(* IEC 61131-3 sources: daoli-st-library/DL_MathData (part 14) *)

(* ---- FC_DL_GearModuleFromCpCalc.st ---- *)
(*
  DL Factory R88 | FC_DL_GearModuleFromCpCalc
  功能：由圆周节 Cp 反算齿轮模数 m=Cp/π，并校验模数是否落在 [min,max] 允许区间
  开源溯源：无（clean-room 自研，依据公开工艺公式 圆周节-模数关系 m=Cp/π，许可证=MIT，借鉴点=公式结构）
  规则：R1-R16 全遵守；R88 简单件标量形（纯标量入参出参，无循环体、无方法、无属性、无数组）
*)
FUNCTION FC_DL_GearModuleFromCpCalc : REAL
VAR_INPUT
    fCpMm : REAL := 12.56637; // 圆周节 Cp（分度圆上相邻同侧齿廓的弧长） [mm] / circular pitch [mm]
    fModuleMin : REAL := 1.0; // 模数允许下限 [mm] / lower allowed module [mm]
    fModuleMax : REAL := 10.0; // 模数允许上限 [mm] / upper allowed module [mm]
END_VAR
VAR_OUTPUT
    fModuleMm : REAL; // 反算模数 m [mm] / back calculated module [mm]
    xInRange : BOOL; // TRUE=模数落在允许区间 [-] / TRUE when module inside the band [-]
END_VAR
VAR
    fPiC : REAL; // 圆周率常数（REAL 精度装入，避免长字面量截断） [-] / pi constant in REAL precision [-]
END_VAR

// 段 1｜出口预置
FC_DL_GearModuleFromCpCalc := -1.0; // 哨兵返回 -1（无效） [-] / sentinel return -1, invalid [-]
fModuleMm := 0.0; // 模数出口预置零 [mm] / module output preset zero [mm]
xInRange := FALSE; // 区间位预置 FALSE（未判定前不认合格） [-] / in-range preset false [-]
fPiC := 3.14159265; // π 常数装入，无量纲 [-] / load the pi constant, dimensionless [-]

// 段 2｜非有限拦截 + 域闸
IF NOT (fCpMm > -1.0E30 AND fCpMm < 1.0E30) OR NOT (fModuleMin > -1.0E30 AND fModuleMin < 1.0E30) OR NOT (fModuleMax > -1.0E30 AND fModuleMax < 1.0E30) THEN
    RETURN; // 三入参任一非有限（NaN/±Inf）即拒算 [-] / any non finite input rejected [-]
END_IF
IF fCpMm < 1.0E-9 THEN
    RETURN; // 周节正域闸：分母 π 恒正，此处拦非正的周节输入 [mm] / positive circular pitch gate [mm]
END_IF
IF fModuleMin < 1.0E-9 OR fModuleMax <= fModuleMin THEN
    RETURN; // 区间自洽闸：下限须为正、上限须严格大于下限 [mm] / band consistency gate [mm]
END_IF

// 段 3｜计算
fModuleMm := fCpMm / fPiC; // mm ÷ 无量纲 = mm，即 m=Cp/π / [mm] / [-] = [mm], m = Cp / pi

// 段 4｜判定与饱和
IF NOT (fModuleMm > -1.0E30 AND fModuleMm < 1.0E30) THEN
    RETURN; // 商结果非有限再拦一次，防溢出成 Inf [-] / re-check the quotient for finiteness [-]
END_IF
xInRange := (fModuleMm >= fModuleMin) AND (fModuleMm <= fModuleMax); // 双侧闭区间直比（含边界） [mm] / closed two sided band compare [mm]

// 段 5｜出口自检
IF fModuleMm < 1.0E-9 THEN
    RETURN; // 出口自检：模数须为正，否则退回哨兵 [mm] / exit self-check, module must be positive [mm]
END_IF
FC_DL_GearModuleFromCpCalc := fModuleMm; // 返回反算模数 [mm] / return the back calculated module [mm]
END_FUNCTION

(* ---- FC_DL_GearRootCircleCalc.st ---- *)
(*
  DL Factory R88 | FC_DL_GearRootCircleCalc
  功能：由模数/齿数算齿根圆直径 df=m(z-2.5)（等价 d-2hf，hf=1.25m），齿数域闸 z>=8
  开源溯源：无（clean-room 自研，依据公开工艺公式 齿根圆直径式 df=m(z-2.5)，许可证=MIT，借鉴点=公式结构）
  规则：R1-R16 全遵守；R88 简单件标量形（纯标量入参出参，无循环体、无方法、无属性、无数组）
*)
FUNCTION FC_DL_GearRootCircleCalc : REAL
VAR_INPUT
    fModuleMm : REAL := 3.0; // 模数 m [mm] / module [mm]
    nTeeth : DINT := 20; // 齿数 z，域闸 z>=8 防齿根自交 [枚] / tooth count, gated at 8 or more [-]
    fDedFactor : REAL := 1.25; // 齿根高系数 hf*=1.25，使 2hf*=2.5 与公式一致 [-] / dedendum coefficient [-]
END_VAR
VAR_OUTPUT
    fDfMm : REAL; // 齿根圆直径 df [mm] / root circle diameter [mm]
    fDedendumMm : REAL; // 齿根高 hf=hf*·m [mm] / dedendum height [mm]
END_VAR
VAR
    fTeeth : REAL; // 齿数实数化结果 [-] / tooth count converted to REAL [-]
    fPitchDiaMm : REAL; // 分度圆直径 d=m·z [mm] / pitch circle diameter [mm]
END_VAR

// 段 1｜出口预置
FC_DL_GearRootCircleCalc := -1.0; // 哨兵返回 -1（无效） [-] / sentinel return -1, invalid [-]
fDfMm := 0.0; // 齿根圆直径预置零 [mm] / root diameter preset zero [mm]
fDedendumMm := 0.0; // 齿根高预置零 [mm] / dedendum preset zero [mm]
fTeeth := 0.0; // 齿数实数预置零 [-] / real teeth preset zero [-]
fPitchDiaMm := 0.0; // 分度圆直径预置零 [mm] / pitch diameter preset zero [mm]

// 段 2｜非有限拦截 + 域闸
IF NOT (fModuleMm > -1.0E30 AND fModuleMm < 1.0E30) OR NOT (fDedFactor > -1.0E30 AND fDedFactor < 1.0E30) THEN
    RETURN; // 模数/齿根高系数任一非有限即拒算 [-] / any non finite input rejected [-]
END_IF
IF fModuleMm < 1.0E-9 THEN
    RETURN; // 模数正域闸 [mm] / positive module gate [mm]
END_IF
IF fDedFactor < 0.8 OR fDedFactor > 1.6 THEN
    RETURN; // 齿根高系数工程域闸（0.8~1.6，标准 1.25） [-] / dedendum coefficient domain gate [-]
END_IF
IF nTeeth < 8 THEN
    RETURN; // 齿数域闸 z>=8：低于 8 齿时齿根圆退化、公式失真 [枚] / root circle degenerates below 8 teeth [-]
END_IF

// 段 3｜计算
fTeeth := DINT_TO_REAL(nTeeth); // DINT→REAL 标准转换函数（R10） [-] / standard conversion function (R10) [-]
fDedendumMm := fDedFactor * fModuleMm; // 无量纲 × mm = mm，hf=hf*·m / [-] × [mm] = [mm]
fPitchDiaMm := fModuleMm * fTeeth; // mm × 无量纲 = mm，d=m·z / [mm] × [-] = [mm]
fDfMm := fPitchDiaMm - 2.0 * fDedendumMm; // mm - mm = mm，df=d-2hf=m(z-2.5) / [mm]

// 段 4｜判定与饱和
IF fDfMm <= 0.0 THEN
    RETURN; // 结果闸：齿根圆直径必须为正，否则齿形无意义 [mm] / root diameter must be positive [mm]
END_IF
IF fDfMm >= fPitchDiaMm THEN
    RETURN; // 结构自洽闸：齿根圆必须小于分度圆 [mm] / structural check df < d [mm]
END_IF

// 段 5｜出口自检
IF NOT (fDfMm > -1.0E30 AND fDfMm < 1.0E30) THEN
    RETURN; // 出口自检：结果非有限即退回哨兵 [mm] / exit self-check on finiteness [mm]
END_IF
FC_DL_GearRootCircleCalc := fDfMm; // 返回齿根圆直径 [mm] / return the root circle diameter [mm]
END_FUNCTION

(* ---- FC_DL_GearSpanMeasurementCalc.st ---- *)
(*
  DL Factory R88 | FC_DL_GearSpanMeasurementCalc
  功能：由模数/齿数/压力角算跨 k 齿公法线长度 Wk=m·cosα·[π(k-0.5)+z·invα]
  开源溯源：无（clean-room 自研，依据公开工艺公式 跨齿公法线长度式，许可证=MIT，借鉴点=公式结构）
  规则：R1-R16 全遵守；R88 简单件标量形（纯标量入参出参，无循环体、无方法、无属性、无数组）
*)
FUNCTION FC_DL_GearSpanMeasurementCalc : REAL
VAR_INPUT
    fModuleMm : REAL := 3.0; // 模数 m [mm] / module [mm]
    nTeeth : DINT := 20; // 齿数 z（整数入参，无 NaN 可能，需 z>=5） [枚] / tooth count [-]
    fPressureDeg : REAL := 20.0; // 分度圆压力角 α（度制，域闸 10~30） [°] / pressure angle in degrees [-]
END_VAR
VAR_OUTPUT
    fWkMm : REAL; // 跨 k 齿公法线长度 Wk [mm] / span measurement over k teeth [mm]
    nSpanTeeth : REAL; // 跨齿数 k（REAL 承载的近似整数） [枚] / number of spanned teeth as a real [-]
END_VAR
VAR
    fTeeth : REAL; // 齿数实数化结果 [-] / tooth count converted to REAL [-]
    fAlphaRad : REAL; // 压力角弧度值 [rad] / pressure angle in radians [rad]
    fInvAlpha : REAL; // 渐开线函数 invα=tanα-α(rad) [rad] / involute function [rad]
    fK : REAL; // 取整后的跨齿数 [枚] / truncated span count [-]
    fCosAlpha : REAL; // 压力角余弦 [-] / cosine of the pressure angle [-]
END_VAR

// 段 1｜出口预置
FC_DL_GearSpanMeasurementCalc := -1.0; // 哨兵返回 -1（无效） [-] / sentinel return -1, invalid [-]
fWkMm := 0.0; // 公法线长度预置零 [mm] / span measurement preset zero [mm]
nSpanTeeth := 0.0; // 跨齿数预置零 [枚] / span teeth preset zero [-]

// 段 2｜非有限拦截 + 域闸
IF NOT (fModuleMm > -1.0E30 AND fModuleMm < 1.0E30) OR NOT (fPressureDeg > -1.0E30 AND fPressureDeg < 1.0E30) THEN
    RETURN; // 模数/压力角任一非有限即拒算 [-] / any non finite input rejected [-]
END_IF
IF fModuleMm < 1.0E-9 THEN
    RETURN; // 模数正域闸 [mm] / positive module gate [mm]
END_IF
IF fPressureDeg <= 10.0 OR fPressureDeg >= 30.0 THEN
    RETURN; // 压力角开区间域闸 (10°,30°)，防 invα 与 k 估算同时失真 [°] / open interval gate on alpha [deg]
END_IF
IF nTeeth < 5 THEN
    RETURN; // 齿数下限闸：z<5 时跨齿数估算式不成立 [枚] / span formula invalid below 5 teeth [-]
END_IF

// 段 3｜计算
fTeeth := DINT_TO_REAL(nTeeth); // DINT→REAL 标准转换函数（R10 禁构造函数式） [-] / standard conversion (R10) [-]
fAlphaRad := fPressureDeg * 0.0174532925; // 度 × (π/180) = rad，换算常数 0.0174532925 [rad] / degrees to radians [rad]
fInvAlpha := TAN(fAlphaRad) - fAlphaRad; // tanα-α 均取弧度，结果弧度制 [rad] / involute function in radians [rad]
fCosAlpha := COS(fAlphaRad); // 无量纲 [-] / dimensionless cosine [-]
// 跨齿数估算：k = ROUND(z·α/180 + 0.5)（标准表 z=20/α=20°→3、z=30→4、z=40→5）；正数下 ROUND 等价 TRUNC(x+1)
fK := TRUNC(fTeeth * fPressureDeg / 180.0 + 1.0); // 数学等价 ROUND(z·α/180+0.5)（R88 修复：原式少 1 齿） [枚] / span count [-]
IF fK < 1.0 THEN
    fK := 1.0; // 饱和：跨齿数至少 1，防 k<=0 使公式失效 [枚] / saturate the span count at one [-]
END_IF
nSpanTeeth := fK; // 跨齿数出口（REAL 承载近似整数） [枚] / export span teeth as a real [-]
fWkMm := fModuleMm * fCosAlpha * (3.14159265 * (fK - 0.5) + fTeeth * fInvAlpha); // mm × [-] × [-] = mm，Wk [mm] / span measurement [mm]
IF fWkMm <= 0.0 THEN
    RETURN; // 结果闸：公法线长度必须为正，否则跨齿数取值失败 [mm] / span length must be positive [mm]
END_IF

// 段 4｜判定与饱和
IF NOT (fWkMm > -1.0E30 AND fWkMm < 1.0E30) THEN
    RETURN; // 结果非有限再拦一次 [-] / re-check the result for finiteness [-]
END_IF

// 段 5｜出口自检
IF nSpanTeeth < 1.0 OR nSpanTeeth >= fTeeth THEN
    RETURN; // 出口自检：跨齿数须在 [1,z) 内，否则出口不自洽 [枚] / span count must lie in [1,z) [-]
END_IF
FC_DL_GearSpanMeasurementCalc := fWkMm; // 返回跨 k 齿公法线长度 [mm] / return the span measurement [mm]
END_FUNCTION

(* ---- FC_DL_GearToothThicknessCalc.st ---- *)
(*
  DL Factory R88 | FC_DL_GearToothThicknessCalc
  功能：由模数/齿数算分度圆弦齿厚 s=m·z·sin(π/(2z))，并给出弧齿厚 πm/2 参考值，齿数域闸 z>=6
  开源溯源：无（clean-room 自研，依据公开工艺公式 分度圆弦齿厚式 s=d·sin(π/2z)，许可证=MIT，借鉴点=公式结构）
  规则：R1-R16 全遵守；R88 简单件标量形（纯标量入参出参，无循环体、无方法、无属性、无数组）
*)
FUNCTION FC_DL_GearToothThicknessCalc : REAL
VAR_INPUT
    fModuleMm : REAL := 3.0; // 模数 m [mm] / module [mm]
    nTeeth : DINT := 20; // 齿数 z，域闸 z>=6 [枚] / tooth count, gated at 6 or more [-]
    fHalfAngleMaxRad : REAL := 1.5; // 半齿角上限保护（π/(2z) 须小于此值，防高齿数误用） [rad] / half tooth angle ceiling [rad]
END_VAR
VAR_OUTPUT
    fChordThkMm : REAL; // 分度圆弦齿厚 s [mm] / chordal tooth thickness [mm]
    fArcThkMm : REAL; // 分度圆弧齿厚 πm/2（参考值） [mm] / circular tooth thickness reference [mm]
END_VAR
VAR
    fTeeth : REAL; // 齿数实数化结果 [-] / tooth count converted to REAL [-]
    fHalfAngleRad : REAL; // 半齿角 π/(2z) [rad] / half tooth angle [rad]
    fDenomTeeth : REAL; // 半齿角分母 2z（除零判据） [枚] / half angle denominator [-]
END_VAR

// 段 1｜出口预置
FC_DL_GearToothThicknessCalc := -1.0; // 哨兵返回 -1（无效） [-] / sentinel return -1, invalid [-]
fChordThkMm := 0.0; // 弦齿厚预置零 [mm] / chordal thickness preset zero [mm]
fArcThkMm := 0.0; // 弧齿厚预置零 [mm] / circular thickness preset zero [mm]
fTeeth := 0.0; // 齿数实数预置零 [-] / real teeth preset zero [-]
fHalfAngleRad := 0.0; // 半齿角预置零 [rad] / half angle preset zero [rad]
fDenomTeeth := 0.0; // 分母预置零 [枚] / denominator preset zero [-]

// 段 2｜非有限拦截 + 域闸
IF NOT (fModuleMm > -1.0E30 AND fModuleMm < 1.0E30) OR NOT (fHalfAngleMaxRad > -1.0E30 AND fHalfAngleMaxRad < 1.0E30) THEN
    RETURN; // 模数/保护限任一非有限即拒算 [-] / any non finite input rejected [-]
END_IF
IF fModuleMm < 1.0E-9 THEN
    RETURN; // 模数正域闸 [mm] / positive module gate [mm]
END_IF
IF fHalfAngleMaxRad <= 0.0 THEN
    RETURN; // 保护限正域闸：须为正，否则后面判据失效 [rad] / positive ceiling gate [rad]
END_IF
IF nTeeth < 6 THEN
    RETURN; // 齿数域闸 z>=6：齿数过低时弦齿厚式与齿形均失真 [枚] / tooth count gate for the chord formula [-]
END_IF

// 段 3｜计算
fTeeth := DINT_TO_REAL(nTeeth); // DINT→REAL 标准转换函数（R10） [-] / standard conversion function (R10) [-]
fDenomTeeth := 2.0 * fTeeth; // 无量纲 × 无量纲 = 无量纲，即 2z [-] / the 2z denominator [-]
IF fDenomTeeth < 1.0E-9 THEN
    RETURN; // 除法前分母闸：2z 必须大于 1E-9 才可作除数 [-] / denominator gate before the division [-]
END_IF
fHalfAngleRad := 3.14159265 / fDenomTeeth; // 无量纲 ÷ 无量纲 = rad，π/(2z) [rad] / half tooth angle [rad]
IF fHalfAngleRad >= fHalfAngleMaxRad THEN
    RETURN; // 半齿角上限闸：超出说明齿数或输入落入误用区间 [rad] / half angle ceiling check [rad]
END_IF
fChordThkMm := fModuleMm * fTeeth * SIN(fHalfAngleRad); // mm × [-] × [-] = mm，s=m·z·sin(π/2z) / [mm]
fArcThkMm := 3.14159265 * fModuleMm * 0.5; // 无量纲 × mm × 0.5 = mm，πm/2（以乘 0.5 替除 2） / [mm]

// 段 4｜判定与饱和
IF fChordThkMm <= 0.0 OR fChordThkMm >= fArcThkMm THEN
    RETURN; // 结构自洽闸：弦齿厚须为正且小于弧齿厚 [mm] / chord thickness must lie in (0, arc) [mm]
END_IF

// 段 5｜出口自检
IF NOT (fChordThkMm > -1.0E30 AND fChordThkMm < 1.0E30) THEN
    RETURN; // 出口自检：结果非有限即退回哨兵 [mm] / exit self-check on finiteness [mm]
END_IF
FC_DL_GearToothThicknessCalc := fChordThkMm; // 返回分度圆弦齿厚 [mm] / return the chordal tooth thickness [mm]
END_FUNCTION

(* ---- FC_DL_GeoBBoxFromPtsFixed.st ---- *)
(*==============================================================================
 * 组件名称 : FC_DL_GeoBBoxFromPtsFixed ｜ 子库 : DL_MathData ｜ v1.0.0 ｜ 2026-11-24
 * 平台     : CODESYS 3.5 / TwinCAT 3 / InoProShop / Machine Expert（纯 IEC，无厂商库）
 * 功能简介 : 定长点列的轴对齐包围盒（BBox）。出参四个极值，用于视觉 ROI 自动贴合、
 *            轨迹占位评估、图形显示自适应缩放。
 * 契约     : 成功返回 TRUE 并写出 fMinX / fMaxX / fMinY / fMaxY；nCnt < 1 时返回 FALSE、
 *            bError := TRUE、四出参置 0；nCnt > 10 时钳到 10 继续（钳位为确定结论）。
 *            数组定长 ARRAY[1..10]，禁变长形参（R17）。
 * 依赖     : 无 DL_ 内部依赖（R16 自足实现），无标准库函数调用
 * 错误码   : R297 零码位范式：eErr 恒 0，仅以 bError / bValid 表达
 * 红线自检 : R1 零全局 R2 零%I/%Q R3 纯IEC R4 点数先钳位后进循环、非有限点跳过并置标志
 *            R5 双语注释 R6 N/A（无状态机）R7 N/A（无定时器/沿实例）
 *            R10 无类型转换 R11 全声明行分号 R15 标识符零保留字冲突
 *            R17 定长数组 R18 N/A（无 bReset）
 * 遗留假设 : 极值初始化取第一个有效点而非 0，避免全正坐标集被 0 拉低下界。
 * 修订历史 : 2026-11-24 R79-A 首版（平面几何族 7/8）
 *============================================================================*)
FUNCTION FC_DL_GeoBBoxFromPtsFixed : BOOL
VAR_INPUT
    aPtsX   : ARRAY[1..10] OF LREAL;    // 点列 X 坐标，1..10 定长 [mm] / X coordinates of the points, fixed length [mm]
    aPtsY   : ARRAY[1..10] OF LREAL;    // 点列 Y 坐标，1..10 定长 [mm] / Y coordinates of the points, fixed length [mm]
    nCnt    : INT;                      // 有效点数，1~10，越界钳位 [个] / effective point count from one to ten, clamped [count]
END_VAR
VAR_OUTPUT
    eErr    : UDINT;    // 错误码，零码位范式恒 0 / error id, always zero under the zero-code rule
    bError  : BOOL;     // 有效点数为零或全为非有限点为真 / TRUE when no usable point exists
    bValid  : BOOL;     // 出参可用标志 / TRUE when the outputs are usable
    fMinX   : LREAL;    // X 下界，故障时 0 [mm] / lower X bound, zero on fault [mm]
    fMaxX   : LREAL;    // X 上界，故障时 0 [mm] / upper X bound, zero on fault [mm]
    fMinY   : LREAL;    // Y 下界，故障时 0 [mm] / lower Y bound, zero on fault [mm]
    fMaxY   : LREAL;    // Y 上界，故障时 0 [mm] / upper Y bound, zero on fault [mm]
END_VAR
VAR CONSTANT
    DL_PTS_MAX : INT := 10;         // 点列定长上限 [个] / fixed capacity of the point arrays [count]
    DL_PTS_MIN : INT := 1;          // 最少有效点数 [个] / minimum usable point count [count]
    DL_ONE     : INT := 1;          // 下标步长与 1 基起始 [个] / index step and the one based start [count]
    DL_FIN_LIM : LREAL := 1.0E308;  // 有限性上界，超过按无穷处置 [mm] / finiteness ceiling [mm]
    DL_ZERO_L  : LREAL := 0.0;      // 实数零哨兵 [mm] / real zero sentinel [mm]
END_VAR
VAR
    nUse    : INT;      // 钳位后的有效点数 [个] / effective point count after clamping [count]
    nSeen   : INT;      // 已纳入极值的有效点数 [个] / points that entered the extremes [count]
    i       : INT;      // 遍历索引，1 起 [个] / loop index starting at one [count]
    fX      : LREAL;    // 当前点 X 快照 [mm] / X snapshot of the current point [mm]
    fY      : LREAL;    // 当前点 Y 快照 [mm] / Y snapshot of the current point [mm]
END_VAR

// 段 1｜出口预置 / segment 1, preset the exit
FC_DL_GeoBBoxFromPtsFixed := FALSE;     // 缺省失败 / default failure
eErr   := 0;                            // 零码位范式 / zero-code rule
bError := FALSE;                        // 预置无故障 / preset no fault
bValid := FALSE;                        // 域闸前不认出参 / the outputs are unusable until the gates pass
fMinX  := DL_ZERO_L;                    // 下界清零 / clear the lower bound
fMaxX  := DL_ZERO_L;                    // 上界清零 / clear the upper bound
fMinY  := DL_ZERO_L;                    // 下界清零 / clear the lower bound
fMaxY  := DL_ZERO_L;                    // 上界清零 / clear the upper bound

// 段 2｜点数钳位与下越界拦截 / segment 2, clamp the count and reject an empty set
nUse := nCnt;
IF nUse > DL_PTS_MAX THEN
    nUse := DL_PTS_MAX;                 // 钳到定长上限 / clamp to the fixed capacity
END_IF
IF nUse < DL_PTS_MIN THEN
    bError := TRUE;                     // 无点可统计 / no point to scan
    RETURN;
END_IF
nSeen := 0;                             // 已纳入点计数清零 / clear the accepted counter

// 段 3｜单趟扫描：首个有效点建立初值，其后逐点更新 / segment 3, one pass with the first usable point as seed
FOR i := DL_ONE TO nUse DO
    fX := aPtsX[i];                     // X 快照 / X snapshot
    fY := aPtsY[i];                     // Y 快照 / Y snapshot
    IF NOT ((fX <> fX) OR (ABS(fX) > DL_FIN_LIM) OR (fY <> fY) OR (ABS(fY) > DL_FIN_LIM)) THEN
        IF nSeen = 0 THEN
            fMinX := fX;                // 首点种子，避免 0 被当极值 / seed from the first point instead of zero
            fMaxX := fX;
            fMinY := fY;
            fMaxY := fY;
        ELSE
            IF fX < fMinX THEN
                fMinX := fX;            // 更新 X 下界 / update the lower X bound
            END_IF
            IF fX > fMaxX THEN
                fMaxX := fX;            // 更新 X 上界 / update the upper X bound
            END_IF
            IF fY < fMinY THEN
                fMinY := fY;            // 更新 Y 下界 / update the lower Y bound
            END_IF
            IF fY > fMaxY THEN
                fMaxY := fY;            // 更新 Y 上界 / update the upper Y bound
            END_IF
        END_IF
        nSeen := nSeen + DL_ONE;        // 有效点计数 / count the accepted point
    END_IF
END_FOR

// 段 4｜出口：全为非有限点按故障处置 / segment 4, exit with the all non finite case treated as a fault
IF nSeen = 0 THEN
    bError := TRUE;                     // 全部点非有限 / every point is non finite
    fMinX  := DL_ZERO_L;                // 出参归零 / zero the outputs
    fMaxX  := DL_ZERO_L;
    fMinY  := DL_ZERO_L;
    fMaxY  := DL_ZERO_L;
    RETURN;
END_IF
bValid := TRUE;                         // 出参可用 / the outputs are usable
FC_DL_GeoBBoxFromPtsFixed := TRUE;      // 求解成功 / the request succeeded
END_FUNCTION

(* ---- FC_DL_GeoCentroid3Pt.st ---- *)
(*==============================================================================
 * 组件名称 : FC_DL_GeoCentroid3Pt ｜ 子库 : DL_MathData ｜ v1.0.0 ｜ 2026-11-24
 * 平台     : CODESYS 3.5 / TwinCAT 3 / InoProShop / Machine Expert（纯 IEC，无厂商库）
 * 功能简介 : 三顶点三角形质心（重心）坐标。出参 fCx = (x1+x2+x3)/3、fCy = (y1+y2+y3)/3。
 *            用于三点示教求工位中心、三点视觉定位求零件中心、夹具三支撑点配平。
 * 契约     : 成功返回 TRUE 并写出质心；三点共线（|叉积| < 1.0E-9）返回 FALSE、
 *            bError := TRUE、出参置 0 —— 共线三角形无质心可言，不得返回中点冒充。
 * 依赖     : 无 DL_ 内部依赖（R16 自足实现）；Standard.library: ABS
 * 错误码   : R297 零码位范式：eErr 恒 0，仅以 bError / bValid 表达
 * 红线自检 : R1 零全局 R2 零%I/%Q R3 纯IEC R4 NaN 自反判据 + 无穷上界 + 共线前拦、
 *            除数为常量 3 ｜ R5 双语注释 R6 N/A（无状态机）R7 N/A（无定时器/沿实例）
 *            R10 无类型转换 R11 全声明行分号 R15 标识符零保留字冲突 R18 N/A（无 bReset）
 * 修订历史 : 2026-11-24 R79-A 首版（平面几何族 5/8）
 *============================================================================*)
FUNCTION FC_DL_GeoCentroid3Pt : BOOL
VAR_INPUT
    fX1     : LREAL;    // 顶点一 X [mm] / X of the first vertex [mm]
    fY1     : LREAL;    // 顶点一 Y [mm] / Y of the first vertex [mm]
    fX2     : LREAL;    // 顶点二 X [mm] / X of the second vertex [mm]
    fY2     : LREAL;    // 顶点二 Y [mm] / Y of the second vertex [mm]
    fX3     : LREAL;    // 顶点三 X [mm] / X of the third vertex [mm]
    fY3     : LREAL;    // 顶点三 Y [mm] / Y of the third vertex [mm]
END_VAR
VAR_OUTPUT
    eErr    : UDINT;    // 错误码，零码位范式恒 0 / error id, always zero under the zero-code rule
    bError  : BOOL;     // 三点共线或输入非有限为真 / TRUE on collinear points or non finite inputs
    bValid  : BOOL;     // 出参可用标志 / TRUE when the outputs are usable
    fCx     : LREAL;    // 质心 X 坐标，故障时 0 [mm] / centroid X, zero on fault [mm]
    fCy     : LREAL;    // 质心 Y 坐标，故障时 0 [mm] / centroid Y, zero on fault [mm]
END_VAR
VAR CONSTANT
    DL_EPS      : LREAL := 1.0E-9;      // 共线判据容差，小于它视为共线 [mm²] / collinearity tolerance [mm²]
    DL_FIN_LIM  : LREAL := 1.0E308;     // 有限性上界 [mm] / finiteness ceiling [mm]
    DL_THREE    : LREAL := 3.0;         // 顶点数，质心的除数 [个] / vertex count, the centroid divisor
    DL_ZERO_L   : LREAL := 0.0;         // 实数零哨兵 / real zero sentinel
END_VAR
VAR
    fCross  : LREAL;    // 两倍有向面积的叉积 [mm²] / cross product, twice the signed area [mm²]
END_VAR

// 段 1｜出口预置 / segment 1, preset the exit
FC_DL_GeoCentroid3Pt := FALSE;      // 缺省失败 / default failure
eErr   := 0;                        // 零码位范式 / zero-code rule
bError := FALSE;                    // 预置无故障 / preset no fault
bValid := FALSE;                    // 域闸前不认出参 / the outputs are unusable until the gates pass
fCx    := DL_ZERO_L;                // 质心 X 清零 / clear the centroid X
fCy    := DL_ZERO_L;                // 质心 Y 清零 / clear the centroid Y

// 段 2｜非有限闸：六个坐标任一为 NaN 即拒 / segment 2, the non finite gate
IF (fX1 <> fX1) OR (fY1 <> fY1) OR (fX2 <> fX2) OR (fY2 <> fY2) OR (fX3 <> fX3) OR (fY3 <> fY3) THEN
    bError := TRUE;                 // 含非数输入 / a not a number input was seen
    RETURN;
END_IF

// 段 3｜共线闸：叉积即两倍有向面积，近零则三点共线 / segment 3, the collinearity gate
fCross := ((fX2 - fX1) * (fY3 - fY1)) - ((fY2 - fY1) * (fX3 - fX1));
IF (fCross <> fCross) OR (ABS(fCross) > DL_FIN_LIM) THEN
    bError := TRUE;                 // 叉积非有限 / the cross product is not finite
    RETURN;
END_IF
IF ABS(fCross) < DL_EPS THEN
    bError := TRUE;                 // 三点共线，无质心 / the points are collinear and no centroid exists
    RETURN;
END_IF

// 段 4｜质心：三坐标算术平均，除数为常量 3 / segment 4, the arithmetic mean of the three vertices
fCx := (fX1 + fX2 + fX3) / DL_THREE;    // 质心 X / centroid X
fCy := (fY1 + fY2 + fY3) / DL_THREE;    // 质心 Y / centroid Y
bValid := TRUE;                         // 出参可用 / the outputs are usable
FC_DL_GeoCentroid3Pt := TRUE;           // 求解成功 / the request succeeded
END_FUNCTION

(* ---- FC_DL_GeoChordHeightCalc.st ---- *)
(*==============================================================================
 * 组件名称 : FC_DL_GeoChordHeightCalc ｜ 子库 : DL_MathData ｜ v1.0.0 ｜ 2026-11-24
 * 平台     : CODESYS 3.5 / TwinCAT 3 / InoProShop / Machine Expert（纯 IEC，无厂商库）
 * 功能简介 : 圆弧弦高（弓高/矢高）h = r − √(r² − (c/2)²)。供圆弧插补弦高误差限、
 *            板材折弯回弹补偿、视觉圆检测圆度评估使用。
 * 契约     : r ≤ 0、c ≤ 0、c > 2r（容差 1.0E-9）、入参非有限 → 返回 0、bError := TRUE、
 *            bValid := FALSE；合法 → 返回 ≥ 0 的弦高、bValid := TRUE。
 * 依赖     : 无 DL_ 内部依赖（R16 自足实现），仅用标准库 SQRT / ABS
 * 错误码   : R297 零码位范式：eErr 恒 0，仅以 bError / bValid 表达
 * 红线自检 : R1 零全局 R2 零%I/%Q R3 纯IEC R4 浮点容差 1.0E-9 + 判别式防负 + 非有限拦截
 *            R5 双语注释 R6 N/A（无状态机）R7 N/A（无定时器/沿实例）
 *            R10 无类型转换 R11 全声明行分号 R15 标识符零保留字冲突
 * 遗留假设 : 弦长等于直径时弦高等于半径（半圆），容差带内的 c 略大于 2r 视为合法并按
 *            判别式归零处理；NaN 用自反判（x <> x），Inf 用自减判（x − x 非零）。
 * 修订历史 : 2026-11-24 R79-B 首版（几何族 1/3）
 *============================================================================*)
FUNCTION FC_DL_GeoChordHeightCalc : LREAL
VAR_INPUT
    fRadius : LREAL := 0.0; // 圆弧半径，须 > 0 [mm] / the arc radius, strictly positive
    fChord  : LREAL := 0.0; // 弦长，须 > 0 且 ≤ 2r [mm] / the chord length, positive and at most the diameter
END_VAR
VAR_OUTPUT
    eErr   : UDINT; // 错误码，零码位范式恒 0 / error id, always zero under the zero-code rule
    bError : BOOL;  // 定义域非法或入参非有限时为真 / TRUE on an invalid domain or a non finite input
    bValid : BOOL;  // 返回值可用标志 / TRUE when the return value is usable
END_VAR
VAR CONSTANT
    DL_ZERO : LREAL := 0.0;      // 实数零哨兵 [mm] / the real zero sentinel
    DL_TWO  : LREAL := 2.0;      // 倍数二，直径与半弦换算 [无量纲] / the factor two used for the diameter and the half chord
    DL_TOL  : LREAL := 1.0E-9;   // 浮点容差（本件唯一比较口径）[无量纲] / the single floating tolerance of this component
END_VAR
VAR
    fHalf  : LREAL; // 半弦长 c/2 [mm] / the half chord length
    fDisc  : LREAL; // 判别式 r² − (c/2)²，防负归零后开方 [mm²] / the discriminant, clamped to zero before the square root
    fDiff  : LREAL; // 非有限检测用的自减量 [无量纲] / the self difference used for the infinity probe
END_VAR

// 段 1｜出口预置 / segment 1, preset the exit
FC_DL_GeoChordHeightCalc := DL_ZERO;  // 缺省零 / default zero
eErr   := 0;                          // 零码位范式 / zero-code rule
bError := FALSE;                      // 预置无故障 / preset no fault
bValid := FALSE;                      // 域闸前不认返回值 / the return value is unusable until the gates pass

// 段 2｜非有限拦截：NaN 自反判，Inf 自减判（Inf − Inf = NaN 使自减表达式不等自身）/ segment 2, the non finite gate
IF (fRadius <> fRadius) OR (fChord <> fChord) THEN
    bError := TRUE;                   // NaN 入参 / a NaN input
    RETURN;                           // 返回 0 / return the preset zero
END_IF
fDiff := fRadius - fRadius;           // 半径自减 / the radius self difference
IF fDiff <> DL_ZERO THEN
    bError := TRUE;                   // 半径非有限（Inf）/ the radius is not finite
    RETURN;                           // 返回 0 / return the preset zero
END_IF
fDiff := fChord - fChord;             // 弦长自减 / the chord self difference
IF fDiff <> DL_ZERO THEN
    bError := TRUE;                   // 弦长非有限（Inf）/ the chord is not finite
    RETURN;                           // 返回 0 / return the preset zero
END_IF

// 段 3｜定义域闸：r > 0、c > 0、c ≤ 2r + 容差 / segment 3, the domain gates
IF fRadius <= DL_ZERO THEN
    bError := TRUE;                   // 半径非正 / the radius is not positive
    RETURN;                           // 返回 0 / return the preset zero
END_IF
IF fChord <= DL_ZERO THEN
    bError := TRUE;                   // 弦长非正 / the chord is not positive
    RETURN;                           // 返回 0 / return the preset zero
END_IF
IF fChord > ((DL_TWO * fRadius) + DL_TOL) THEN
    bError := TRUE;                   // 弦长超过直径 / the chord exceeds the diameter
    RETURN;                           // 返回 0 / return the preset zero
END_IF

// 段 4｜判别式防负：容差带内 c 略大于 2r 时 r² − (c/2)² 可能为极小负值，归零后开方 / segment 4, the discriminant clamp
fHalf := fChord / DL_TWO;             // 半弦 [mm] / the half chord
fDisc := (fRadius * fRadius) - (fHalf * fHalf);  // 判别式 [mm²] / the discriminant
IF fDisc < DL_ZERO THEN fDisc := DL_ZERO; END_IF  // 防负归零，避免 SQRT 得 NaN / clamp to zero so the square root stays real

// 段 5｜弦高出口 / segment 5, the sagitta
FC_DL_GeoChordHeightCalc := fRadius - SQRT(fDisc);  // h = r − √(r² − (c/2)²) [mm] / the sagitta
bValid := TRUE;                                     // 返回值可用 / the return value is usable
END_FUNCTION

(* ---- FC_DL_GeoCircleSectorArea.st ---- *)
(*==============================================================================
 * 组件名称 : FC_DL_GeoCircleSectorArea ｜ 子库 : DL_MathData ｜ v1.0.1 ｜ 2026-11-24
 * 平台     : CODESYS 3.5 / TwinCAT 3 / InoProShop / Machine Expert（纯 IEC，无厂商库）
 * 功能简介 : 圆扇形面积 A = 0.5 · r² · θ(rad)。供扇形料片下料、回转台扫掠面积、
 *            风扇扇区通流面积等调用方。角度先按 360 取模归一到 [0,360)，再内联 π/180 转弧度。
 * 契约     : r ≥ 0 且角度有限 → 返回面积、bValid := TRUE（r = 0 合法，面积 0）；
 *            r < 0 或入参非有限 → 返回 0、bError := TRUE、bValid := FALSE。
 * 依赖     : 无 DL_ 内部依赖（R16 自足实现：π 与度弧换算内联，不调用任何换算件）
 * 错误码   : R297 零码位范式：eErr 恒 0，仅以 bError / bValid 表达
 * 红线自检 : R1 零全局 R2 零%I/%Q R3 纯IEC R4 无除法风险（除数恒 360 与 180）+ 非有限拦截
 *            R5 双语注释 R6 N/A（无状态机）R7 N/A（无定时器/沿实例）
 *            R10 无类型转换（取整用 TRUNC 泛型，保持 LREAL）R11 全声明行分号
 *            R15 标识符零保留字冲突
 * 遗留假设 : 取模用「TRUNC(θ/360) 后减整圈」实现在 LREAL 域完成，避免 LREAL_TO_DINT
 *            在大角度下的截断溢出；|θ| 超过 1E15 度时整圈数已超出 LREAL 尾数精度，
 *            余角精度下降（工程角度远小于该量级，故不设上限拦截）；
 *            π 取 3.141592653589793（LREAL 双精度 15~16 位有效数字口径）。
 * 修订历史 : 2026-11-24 R79-B 首版（几何族 2/3）
 *============================================================================*)
FUNCTION FC_DL_GeoCircleSectorArea : LREAL
VAR_INPUT
    fRadius   : LREAL := 0.0; // 圆半径，须 ≥ 0 [mm] / the circle radius, zero allowed
    fAngleDeg : LREAL := 0.0; // 扇区圆心角，可负，内部按 360 取模 [度] / the central angle, negative allowed, wrapped by 360
END_VAR
VAR_OUTPUT
    eErr   : UDINT; // 错误码，零码位范式恒 0 / error id, always zero under the zero-code rule
    bError : BOOL;  // 半径非法或入参非有限时为真 / TRUE on a negative radius or a non finite input
    bValid : BOOL;  // 返回值可用标志 / TRUE when the return value is usable
END_VAR
VAR CONSTANT
    DL_FIN     : LREAL := 1.0E30;  // 有限性判据上界（R477 范式：ABS(x)>FIN 判 Inf，禁用 x-x 差判）/ finiteness ceiling, ABS(x)>FIN flags Inf
    DL_ZERO : LREAL := 0.0;               // 实数零哨兵 [mm] / the real zero sentinel
    DL_HALF : LREAL := 0.5;               // 扇形系数 1/2 [无量纲] / the sector coefficient one half
    DL_FULL : LREAL := 360.0;             // 整圆角度 [度] / the full turn in degrees
    DL_DEG  : LREAL := 180.0;             // 半圆角度，度弧换算分母 [度] / the half turn, the degree to radian divisor
    DL_PI   : LREAL := 3.141592653589793; // 圆周率（内联，不引用换算件）[无量纲] / the inline constant pi
END_VAR
VAR
    fTurns : LREAL; // 整圈数（向零截断，LREAL 域内）[圈] / the whole turn count truncated toward zero
    fAng   : LREAL; // 归一后的圆心角，落在 [0,360) [度] / the wrapped central angle inside one turn
    fRad   : LREAL; // 圆心角弧度值 [弧度] / the central angle in radians
END_VAR

// 段 1｜出口预置 / segment 1, preset the exit
FC_DL_GeoCircleSectorArea := DL_ZERO;  // 缺省零 / default zero
eErr   := 0;                           // 零码位范式 / zero-code rule
bError := FALSE;                       // 预置无故障 / preset no fault
bValid := FALSE;                       // 域闸前不认返回值 / the return value is unusable until the gates pass

// 段 2｜非有限拦截：NaN 自反判，Inf 自减判 / segment 2, the non finite gate
IF (fRadius <> fRadius) OR (fAngleDeg <> fAngleDeg) THEN
    bError := TRUE;                    // NaN 入参 / a NaN input
    RETURN;                            // 返回 0 / return the preset zero
END_IF
IF (ABS(fRadius) > DL_FIN) OR (ABS(fAngleDeg) > DL_FIN) THEN
    bError := TRUE;                    // Inf 入参 / an infinite input
    RETURN;                            // 返回 0 / return the preset zero
END_IF

// 段 3｜半径域闸：负半径无几何意义，零半径面积为零属合法 / segment 3, the radius gate
IF fRadius < DL_ZERO THEN
    bError := TRUE;                    // 负半径 / a negative radius
    RETURN;                            // 返回 0 / return the preset zero
END_IF

// 段 4｜角度归一：θ − TRUNC(θ/360) × 360 落在 (−360, 360)，负向再补一圈到 [0,360) / segment 4, the angle wrap
fTurns := TRUNC(fAngleDeg / DL_FULL);          // 整圈数，向零截断 [圈] / whole turns truncated toward zero
fAng   := fAngleDeg - (fTurns * DL_FULL);      // 余角，与输入同号 [度] / the remainder carrying the input sign
IF fAng < DL_ZERO THEN fAng := fAng + DL_FULL; END_IF  // 负向补一圈 / add one turn for negative remainders

// 段 5｜度转弧度并求面积：A = 0.5 · r² · θ·π/180 / segment 5, the area
fRad := fAng * (DL_PI / DL_DEG);               // 弧度值 [弧度] / the radian value
FC_DL_GeoCircleSectorArea := DL_HALF * fRadius * fRadius * fRad;  // 面积 [mm²] / the sector area
bValid := TRUE;                                // 返回值可用 / the return value is usable
END_FUNCTION

(* ---- FC_DL_GeoLineAngleXY.st ---- *)
(*==============================================================================
 * 组件名称 : FC_DL_GeoLineAngleXY ｜ 子库 : DL_MathData ｜ v1.0.0 ｜ 2026-11-24
 * 平台     : CODESYS 3.5 / TwinCAT 3 / InoProShop / Machine Expert（纯 IEC，无厂商库）
 * 功能简介 : 两点连线相对 X 轴的有向角 [rad]，域 (−π, π]。实现取 ATAN(dy/dx) 加象限补偿，
 *            刻意不用 ATAN2 —— ATAN2 的形参序（先 x 后 y 还是先 y 后 x）在 CODESYS 手册、
 *            TwinCAT 与标准桩之间互不相同，跨平台移植时必出错；ATAN 单形参无此歧义。
 * 契约     : 返回有向角 ∈ (−π, π]；两点重合（距离 < 1.0E-9）返回 0、bError := TRUE、
 *            bValid := FALSE；输入含 NaN 或非有限值时同样按故障处置。
 * 依赖     : 无 DL_ 内部依赖（R16 自足实现）；Standard.library: ATAN / ABS
 * 错误码   : R297 零码位范式：eErr 恒 0，仅以 bError / bValid 表达
 * 红线自检 : R1 零全局 R2 零%I/%Q R3 纯IEC R4 NaN 自反判据 + 无穷上界 + 竖直线单列
 *            （除法前判 dx 容差）｜ R5 双语注释 R6 N/A（无状态机）
 *            R7 N/A（无定时器/沿实例）R10 无类型转换 R11 全声明行分号
 *            R15 标识符零保留字冲突 R18 N/A（无 bReset）
 * 遗留假设 : 象限补偿四分支已覆盖 dx<0 的两种情形与 dx 近零的两种竖直方向，
 *            dx>0 时 ATAN 值本身即落在 (−π/2, π/2)，无需补偿。
 * 修订历史 : 2026-11-24 R79-A 首版（平面几何族 8/8）
 *============================================================================*)
FUNCTION FC_DL_GeoLineAngleXY : LREAL
VAR_INPUT
    fAx     : LREAL;    // 起点 X 坐标 [mm] / X coordinate of the start point [mm]
    fAy     : LREAL;    // 起点 Y 坐标 [mm] / Y coordinate of the start point [mm]
    fBx     : LREAL;    // 终点 X 坐标 [mm] / X coordinate of the end point [mm]
    fBy     : LREAL;    // 终点 Y 坐标 [mm] / Y coordinate of the end point [mm]
END_VAR
VAR_OUTPUT
    eErr    : UDINT;    // 错误码，零码位范式恒 0 / error id, always zero under the zero-code rule
    bError  : BOOL;     // 两点重合或输入非有限为真 / TRUE on coincident points or non finite inputs
    bValid  : BOOL;     // 结果可用标志 / result usable flag
END_VAR
VAR CONSTANT
    DL_EPS      : LREAL := 1.0E-9;                  // 长度容差，短于此值判重合 [mm] / length tolerance for the coincident test [mm]
    DL_FIN_LIM  : LREAL := 1.0E308;                 // 有限性上界 [mm] / finiteness ceiling [mm]
    DL_PI       : LREAL := 3.14159265358979323846;  // 圆周率 [rad] / pi in radians [rad]
    DL_PI_HALF  : LREAL := 1.57079632679489661923;  // 半圆周率，竖直方向角 [rad] / half pi, the vertical angle [rad]
    DL_ZERO_L   : LREAL := 0.0;                     // 实数零哨兵 / real zero sentinel
END_VAR
VAR
    fDx     : LREAL;    // X 方向的增量 [mm] / increment along X [mm]
    fDy     : LREAL;    // Y 方向的增量 [mm] / increment along Y [mm]
    fAng    : LREAL;    // 角度中间量 [rad] / angle interim value [rad]
END_VAR

// 段 1｜出口预置 / segment 1, preset the exit
FC_DL_GeoLineAngleXY := DL_ZERO_L;  // 缺省角 0 / default angle zero
eErr   := 0;                        // 零码位范式 / zero-code rule
bError := FALSE;                    // 预置无故障 / preset no fault
bValid := FALSE;                    // 解算完成前不认结果 / unusable until the solve ends

// 段 2｜非有限闸：四个坐标任一为 NaN 即拒 / segment 2, the non finite gate
IF (fAx <> fAx) OR (fAy <> fAy) OR (fBx <> fBx) OR (fBy <> fBy) THEN
    bError := TRUE;                 // 含非数输入 / a not a number input was seen
    RETURN;
END_IF

// 段 3｜增量与重合判定：两点重合时角度无定义 / segment 3, the increments and the coincident test
fDx := fBx - fAx;
fDy := fBy - fAy;
IF (ABS(fDx) > DL_FIN_LIM) OR (ABS(fDy) > DL_FIN_LIM) THEN
    bError := TRUE;                 // 增量非有限 / the increments are not finite
    RETURN;
END_IF
IF (ABS(fDx) < DL_EPS) AND (ABS(fDy) < DL_EPS) THEN
    bError := TRUE;                 // 两点重合，方向无定义 / the points coincide and no direction exists
    RETURN;
END_IF

// 段 4｜竖直方向单列：dx 近零时角为 ±π/2，避免除以近零量放大误差 / segment 4, the vertical branches
IF ABS(fDx) < DL_EPS THEN
    IF fDy > DL_ZERO_L THEN
        FC_DL_GeoLineAngleXY := DL_PI_HALF;     // 正上方 90° / straight up
    ELSE
        FC_DL_GeoLineAngleXY := -DL_PI_HALF;    // 正下方 −90° / straight down
    END_IF
    bValid := TRUE;                 // 结果可用 / the result is usable
    RETURN;
END_IF

// 段 5｜象限补偿：dx<0 时 ATAN 值需平移 ±π 才能落回 (−π, π] / segment 5, the quadrant compensation
fAng := ATAN(fDy / fDx);            // 主值域 (−π/2, π/2)，除数为已证非零的 dx / principal value with a proven non zero divisor
IF fDx < DL_ZERO_L THEN
    IF fDy > DL_ZERO_L THEN
        fAng := fAng + DL_PI;       // 第二象限 / the second quadrant
    ELSE
        fAng := fAng - DL_PI;       // 第三象限，含 dy = 0 时取 −π 再归到 +π 的边界 / the third quadrant
        IF ABS(fAng) > (DL_PI - DL_EPS) THEN
            fAng := DL_PI;          // 负 X 轴归一到 +π，保证值域 (−π, π] / the negative X axis normalises to plus pi
        END_IF
    END_IF
END_IF

// 段 6｜出口 / segment 6, exit
FC_DL_GeoLineAngleXY := fAng;       // 有向角 [rad] / the signed angle in radians
bValid := TRUE;                     // 结果可用 / the result is usable
END_FUNCTION

(* ---- FC_DL_GeoMeanCalc.st ---- *)
(*==============================================================================
 * 组件名称 (Component)  : FC_DL_GeoMeanCalc
 * 所属子库 (Sublibrary) : DL_MathData
 * 当前版本 (Version)    : 1.0.0
 * 兼容性 (Platform)     : CODESYS 3.5+ / TwinCAT 3 / 汇川 InoProShop / 施耐德 Machine Expert
 *                         仅用标准函数 LN / EXP / ABS，零厂商私有库
 * 功能描述 (Function)   : 非负数组几何平均叶子件。在 log 域求和：g = exp(Σln(xi)/n)，
 *                         避免直接连乘的上溢/下溢（n 件 0.5 连乘即沉到下溢）。
 *                         良率均值、轴承寿命均值、稀释比均值等乘性量场景。
 * 来源标签 (Origin)     : 自研线（IEC 61131-3 标准语义的道莅防御性实现，clean-room）
 * 边界语义 (Boundary)   : ① 拒算闸：任一元素 xi <= eps 或 NaN → bValid = FALSE 且
 *                         返回 0.0（几何平均对非正元素无定义，静默取绝对值会把
 *                         「负良率」这种数据事故伪装成正常结果）；bValid 报告
 *                         拒算，调用方据此走数据质量链而非数值链；
 *                         ② 计数钳位：nCount < 1 → 拒算；nCount > 常量上限 →
 *                         钳位到上限（防越界，R308 口径）；
 *                         ③ ln 域结果超出 exp 可表域时拒绝：Σln/n > 709（LREAL
 *                         exp 上限 ln(1.8E308)≈709.78）→ 拒算防 Inf；
 *                         ④ 纯函数：无状态、无定时器、无副作用。
 * 码位     (Codes)      : 按 R297 范式零 16# 码位硬编码，拒算语义经 bValid 布尔出口承载
 * 红线自检 (Redline)    : 7 项红线已自检：R1 零全局 ✓｜R2 零物理地址 ✓｜R3 纯 IEC ✓
 *                         R4 防御完整（拒算/钳位/exp 域闸/NaN 自反判）✓
 *                         R5 双语同行注释 ✓｜R6 N/A（纯函数无状态机）✓｜R7 N/A（无实例）✓
 * 验收向量 (Acceptance) : V1 输入 [4, 16] → g = 8.0（容差 1E-6）；
 *                         V2 输入含 0 或负数 → bValid = FALSE 返回 0.0；
 *                         V3 nCount = 0 → bValid = FALSE；
 *                         V4 输入 [1,1,1] → g = 1.0（ln 域零和恒等式）。
 * 修订历史 (Revision)   : 2026-11-20  v1.0.0  R49 首版（批 1 · 序号 2）
 *==============================================================================*)
FUNCTION FC_DL_GeoMeanCalc : LREAL           (* 返回几何平均值，拒算路径返回 0.0 / Returns geometric mean, 0.0 on rejection *)
VAR_INPUT
    aVals    : ARRAY[1..32] OF LREAL;        (* 输入数值数组（log 域求和源）[工程单位] / Input value array *)
    nCount   : INT;                          (* 有效元素个数，域 1..32，越界钳位 [件] / Valid element count, clamped to 1..32 *)
END_VAR
VAR_OUTPUT
    bValid   : BOOL;                         (* 本次计算有效性，FALSE = 拒算（含非正元素/计数非法/exp 域溢出）[-] / Validity flag, FALSE = rejected *)
    nRejectReason : INT;                     (* 拒算原因 0 无 1 计数非法 2 非正元素 3 exp 域溢出 [-] / Reject reason code *)
END_VAR
VAR
    i        : INT;                          (* 循环游标（每趟显式初始化，R227）[-] / Loop cursor *)
    nEff     : INT;                          (* 钳位后生效计数 [件] / Clamped effective count *)
    fSumLn   : LREAL;                        (* ln 域累计和 [ln·工程单位] / Accumulated log-domain sum *)
    fMeanLn  : LREAL;                        (* ln 域均值 = fSumLn / n [ln·工程单位] / Log-domain mean *)
    fXi      : LREAL;                        (* 当前元素缓存（防双重下标取值）[工程单位] / Current element cache *)
END_VAR
VAR CONSTANT
    DL_GM_EPS    : LREAL := 1.0E-12;         (* 元素非正判零容差（log 定义域下界）[工程单位] / Non-positive epsilon *)
    DL_GM_LN_MAX : LREAL := 709.0;           (* LREAL 的 exp 可表域上限 [ln] / exp-representable upper bound for LREAL *)
    DL_GM_NMAX   : INT   := 32;              (* 数组容量上限（计数钳位目标）[件] / Array capacity limit *)
END_VAR

(* —— 段 1：缺省输出（R285 全路径赋值） —— *)
FC_DL_GeoMeanCalc := 0.0;                    (* 缺省返回 0.0：可辨识零，不冒充正常结果 / Default 0.0, recognizable zero *)
bValid := FALSE;                             (* 有效性缺省 FALSE / Validity default FALSE *)
nRejectReason := 0;                          (* 拒算原因缺省无 / Reject reason default none *)

(* —— 段 2：计数闸与钳位（下界拒算、上界钳位防数组越界） —— *)
IF nCount < 1 THEN                           (* 零/负计数无统计意义 / Non-positive count meaningless *)
    nRejectReason := 1;                      (* 原因 1：计数非法 / Reason 1: illegal count *)
    RETURN;
END_IF
nEff := nCount;                              (* 生效计数初值 / Effective count init *)
IF nEff > DL_GM_NMAX THEN
    nEff := DL_GM_NMAX;                      (* 计数超容量钳位到上限（R308） / Clamp count to capacity *)
END_IF

(* —— 段 3：逐元素非正闸 + log 域累加（FOR 正步进，可移植） —— *)
FOR i := 1 TO nEff DO
    fXi := aVals[i];                         (* 取当前元素 / Fetch current element *)
    IF (fXi <> fXi) OR (fXi <= DL_GM_EPS) OR ((fXi - fXi) <> (fXi - fXi)) THEN
        nRejectReason := 2;                  (* 原因 2：NaN 或非正元素拒算 / Reason 2: NaN or non-positive rejected *)
        RETURN;                              (* 任一元素非法即整体拒算，不做部分结果 / Whole-call rejection, no partial result *)
    END_IF
    fSumLn := fSumLn + LN(fXi);              (* log 域累加，天然防连乘溢出 / Log-domain accumulation, overflow-free *)
END_FOR

(* —— 段 4：均值与 exp 域闸（除子 = 钳位后计数，恒 >= 1，无除零） —— *)
fMeanLn := fSumLn / INT_TO_LREAL(nCount);    (* ln 域均值，计数已 >= 1（INT_TO_LREAL 显式展宽） / Log-domain mean, explicit widening *)
IF fMeanLn > DL_GM_LN_MAX OR fMeanLn < (-DL_GM_LN_MAX) THEN
    nRejectReason := 3;                      (* 原因 3：exp 域外，防 Inf（R133 非有限值闸前置） / Reason 3: outside exp domain, prevents Inf *)
    RETURN;
END_IF
FC_DL_GeoMeanCalc := EXP(fMeanLn);           (* log 域还原为几何平均 / Exponentiate back to geometric mean *)
bValid := TRUE;                              (* 全闸通过，结果有效 / All gates passed, valid *)
END_FUNCTION

(* ---- FC_DL_GeoPointInConvexQuadXY.st ---- *)
(*==============================================================================
 * 组件名称 : FC_DL_GeoPointInConvexQuadXY ｜ 子库 : DL_MathData ｜ v1.0.0 ｜ 2026-11-24
 * 平台     : CODESYS 3.5 / TwinCAT 3 / InoProShop / Machine Expert（纯 IEC，无厂商库）
 * 功能简介 : 点是否落在凸四边形内（含边界）。顶点须按序（顺或逆时针）给出，
 *            用叉积同号法：点对四条有向边的叉积若全同号（或全近零）即在内部。
 *            用于相机视野分区、机器人安全区、视觉 ROI 的旋转框判定。
 * 契约     : 在内返回 TRUE；四边形退化（|鞋带面积| < 1.0E-6）返回 FALSE、bError := TRUE；
 *            点恰在边上按「在内」处理（容差 1.0E-9）。
 * 依赖     : 无 DL_ 内部依赖（R16 自足实现）；Standard.library: ABS
 * 错误码   : R297 零码位范式：eErr 恒 0，仅以 bError / bValid 表达
 * 红线自检 : R1 零全局 R2 零%I/%Q R3 纯IEC R4 NaN 自反判据 + 无穷上界 + 退化面积极小判据、
 *            浮点无等号判等 ｜ R5 双语注释 R6 N/A（无状态机）R7 N/A（无定时器/沿实例）
 *            R10 无类型转换 R11 全声明行分号 R15 标识符零保留字冲突 R18 N/A（无 bReset）
 * 遗留假设 : 顶点序错乱（如 1-3-2-4）会让叉积法失效并可能误判在外 —— 顶点序由调用方保证，
 *            函数内不做自交检测（自交检测为另件职责）。
 * 修订历史 : 2026-11-24 R79-A 首版（平面几何族 4/8）
 *============================================================================*)
FUNCTION FC_DL_GeoPointInConvexQuadXY : BOOL
VAR_INPUT
    fPx     : LREAL;    // 被测点 X 坐标 [mm] / X coordinate of the measured point [mm]
    fPy     : LREAL;    // 被测点 Y 坐标 [mm] / Y coordinate of the measured point [mm]
    fX1     : LREAL;    // 顶点一 X [mm] / X of the first vertex [mm]
    fY1     : LREAL;    // 顶点一 Y [mm] / Y of the first vertex [mm]
    fX2     : LREAL;    // 顶点二 X [mm] / X of the second vertex [mm]
    fY2     : LREAL;    // 顶点二 Y [mm] / Y of the second vertex [mm]
    fX3     : LREAL;    // 顶点三 X [mm] / X of the third vertex [mm]
    fY3     : LREAL;    // 顶点三 Y [mm] / Y of the third vertex [mm]
    fX4     : LREAL;    // 顶点四 X [mm] / X of the fourth vertex [mm]
    fY4     : LREAL;    // 顶点四 Y [mm] / Y of the fourth vertex [mm]
END_VAR
VAR_OUTPUT
    eErr    : UDINT;    // 错误码，零码位范式恒 0 / error id, always zero under the zero-code rule
    bError  : BOOL;     // 退化四边形或非有限输入为真 / TRUE on a degenerate quad or non finite inputs
    bValid  : BOOL;     // 判定可用标志 / TRUE when the verdict is usable
END_VAR
VAR CONSTANT
    DL_EPS      : LREAL := 1.0E-9;      // 叉积容差，边上的点按「在内」处理 [mm²] / cross tolerance, edge points count as inside [mm²]
    DL_AREA_MIN : LREAL := 1.0E-6;      // 四边形面积下限，小于它判退化 [mm²] / degenerate area threshold [mm²]
    DL_FIN_LIM  : LREAL := 1.0E308;     // 有限性上界 [mm] / finiteness ceiling [mm]
    DL_TWO      : LREAL := 2.0;         // 鞋带面积的二分之一换算 [无量纲] / halving factor of the shoelace sum
END_VAR
VAR
    fArea2  : LREAL;    // 鞋带和，等于两倍面积 [mm²] / shoelace sum, twice the area [mm²]
    fC1     : LREAL;    // 边 1→2 对点的叉积 [mm²] / cross product of edge one to two [mm²]
    fC2     : LREAL;    // 边 2→3 对点的叉积 [mm²] / cross product of edge two to three [mm²]
    fC3     : LREAL;    // 边 3→4 对点的叉积 [mm²] / cross product of edge three to four [mm²]
    fC4     : LREAL;    // 边 4→1 对点的叉积 [mm²] / cross product of edge four to one [mm²]
    bPos    : BOOL;     // 四条叉积是否全为正 / TRUE when every cross product is positive
    bNeg    : BOOL;     // 四条叉积是否全为负 / TRUE when every cross product is negative
END_VAR

// 段 1｜出口预置 / segment 1, preset the exit
FC_DL_GeoPointInConvexQuadXY := FALSE;  // 缺省不在四边形内 / default outside
eErr   := 0;                            // 零码位范式 / zero-code rule
bError := FALSE;                        // 预置无故障 / preset no fault
bValid := FALSE;                        // 判定完成前不可用 / unusable until the verdict ends

// 段 2｜非有限闸：十个坐标任一为 NaN 即拒 / segment 2, the non finite gate
IF (fPx <> fPx) OR (fPy <> fPy) OR (fX1 <> fX1) OR (fY1 <> fY1) OR (fX2 <> fX2) OR (fY2 <> fY2) OR (fX3 <> fX3) OR (fY3 <> fY3) OR (fX4 <> fX4) OR (fY4 <> fY4) THEN
    bError := TRUE;                     // 含非数输入 / a not a number input was seen
    RETURN;
END_IF

// 段 3｜退化闸：鞋带公式求两倍面积，过小即判退化 / segment 3, the shoelace area and the degenerate gate
fArea2 := ABS((fX1 * (fY2 - fY4)) + (fX2 * (fY3 - fY1)) + (fX3 * (fY4 - fY2)) + (fX4 * (fY1 - fY3)));
IF (fArea2 <> fArea2) OR (fArea2 > DL_FIN_LIM) THEN
    bError := TRUE;                     // 面积非有限 / the area is not finite
    RETURN;
END_IF
IF (fArea2 / DL_TWO) < DL_AREA_MIN THEN
    bError := TRUE;                     // 四边形退化（三点共线或重合）/ the quad degenerates
    RETURN;
END_IF

// 段 4｜四条边的叉积：点对每条有向边的相对位置 / segment 4, the four edge cross products
fC1 := ((fX2 - fX1) * (fPy - fY1)) - ((fY2 - fY1) * (fPx - fX1));   // 边 1→2 / edge one to two
fC2 := ((fX3 - fX2) * (fPy - fY2)) - ((fY3 - fY2) * (fPx - fX2));   // 边 2→3 / edge two to three
fC3 := ((fX4 - fX3) * (fPy - fY3)) - ((fY4 - fY3) * (fPx - fX3));   // 边 3→4 / edge three to four
fC4 := ((fX1 - fX4) * (fPy - fY4)) - ((fY1 - fY4) * (fPx - fX4));   // 边 4→1 / edge four to one

// 段 5｜同号判定：全正或全负（近零点按同号处理）/ segment 5, the same sign verdict
bPos := (fC1 > -DL_EPS) AND (fC2 > -DL_EPS) AND (fC3 > -DL_EPS) AND (fC4 > -DL_EPS);
bNeg := (fC1 < DL_EPS) AND (fC2 < DL_EPS) AND (fC3 < DL_EPS) AND (fC4 < DL_EPS);
IF bPos OR bNeg THEN
    FC_DL_GeoPointInConvexQuadXY := TRUE;   // 叉积同号即在凸四边形内 / same signed crosses mean inside
END_IF
bValid := TRUE;                             // 判定可用 / the verdict is usable
END_FUNCTION

(* ---- FC_DL_GeoPointInRectXY.st ---- *)
(*==============================================================================
 * 组件名称 : FC_DL_GeoPointInRectXY ｜ 子库 : DL_MathData ｜ v1.0.0 ｜ 2026-11-24
 * 平台     : CODESYS 3.5 / TwinCAT 3 / InoProShop / Machine Expert（纯 IEC，无厂商库）
 * 功能简介 : 点是否落在轴对齐矩形内（含边界，容差 1.0E-9）。矩形以任意两个对角顶点给出，
 *            宽或高为负时自动换序归一 —— 现场示教常把左上与右下顺序录反，
 *            本件保证录入顺序不影响判定。
 * 契约     : 在内返回 TRUE；任一点含非有限值或矩形退化（宽高均小于容差）时返回 FALSE、
 *            bError := TRUE。边界点按「含」处理（外扩容差）。
 * 依赖     : 无 DL_ 内部依赖（R16 自足实现）；Standard.library: ABS / MIN / MAX
 * 错误码   : R297 零码位范式：eErr 恒 0，仅以 bError / bValid 表达
 * 红线自检 : R1 零全局 R2 零%I/%Q R3 纯IEC R4 NaN 自反判据、浮点无等号判等（全部走容差窗口）
 *            R5 双语注释 R6 N/A（无状态机）R7 N/A（无定时器/沿实例）
 *            R10 无类型转换 R11 全声明行分号 R15 标识符零保留字冲突 R18 N/A（无 bReset）
 * 遗留假设 : 矩形必须轴对齐；旋转框请改用 FC_DL_GeoPointInConvexQuadXY（四边形叉积法）。
 * 修订历史 : 2026-11-24 R79-A 首版（平面几何族 3/8）
 *============================================================================*)
FUNCTION FC_DL_GeoPointInRectXY : BOOL
VAR_INPUT
    fPx     : LREAL;    // 被测点 X 坐标 [mm] / X coordinate of the measured point [mm]
    fPy     : LREAL;    // 被测点 Y 坐标 [mm] / Y coordinate of the measured point [mm]
    fX1     : LREAL;    // 对角顶点一 X，可为大值或小值 [mm] / X of the first corner, may be the larger one [mm]
    fY1     : LREAL;    // 对角顶点一 Y，可为大值或小值 [mm] / Y of the first corner, may be the larger one [mm]
    fX2     : LREAL;    // 对角顶点二 X，可与顶点一顺序任意 [mm] / X of the second corner, order free [mm]
    fY2     : LREAL;    // 对角顶点二 Y，可与顶点一顺序任意 [mm] / Y of the second corner, order free [mm]
END_VAR
VAR_OUTPUT
    eErr    : UDINT;    // 错误码，零码位范式恒 0 / error id, always zero under the zero-code rule
    bError  : BOOL;     // 非有限输入或矩形退化为真 / TRUE on non finite inputs or a degenerate rectangle
    bValid  : BOOL;     // 判定可用标志 / TRUE when the verdict is usable
END_VAR
VAR CONSTANT
    DL_EPS      : LREAL := 1.0E-9;      // 边界容差，边界点按「在内」处理 [mm] / boundary tolerance, edge points count as inside [mm]
    DL_FIN_LIM  : LREAL := 1.0E308;     // 有限性上界 [mm] / finiteness ceiling [mm]
END_VAR
VAR
    fMinX   : LREAL;    // 归一后的 X 下界 [mm] / normalised lower X bound [mm]
    fMaxX   : LREAL;    // 归一后的 X 上界 [mm] / normalised upper X bound [mm]
    fMinY   : LREAL;    // 归一后的 Y 下界 [mm] / normalised lower Y bound [mm]
    fMaxY   : LREAL;    // 归一后的 Y 上界 [mm] / normalised upper Y bound [mm]
END_VAR

// 段 1｜出口预置 / segment 1, preset the exit
FC_DL_GeoPointInRectXY := FALSE;    // 缺省不在矩形内 / default outside
eErr   := 0;                        // 零码位范式 / zero-code rule
bError := FALSE;                    // 预置无故障 / preset no fault
bValid := FALSE;                    // 判定完成前不可用 / unusable until the verdict ends

// 段 2｜非有限闸与量级闸：六个坐标任一为 NaN 或超上界即拒 / segment 2, the non finite and magnitude gates
IF (fPx <> fPx) OR (fPy <> fPy) OR (fX1 <> fX1) OR (fY1 <> fY1) OR (fX2 <> fX2) OR (fY2 <> fY2) THEN
    bError := TRUE;                 // 含非数输入 / a not a number input was seen
    RETURN;
END_IF
IF (ABS(fPx) > DL_FIN_LIM) OR (ABS(fPy) > DL_FIN_LIM) OR (ABS(fX1) > DL_FIN_LIM) OR (ABS(fY1) > DL_FIN_LIM) OR (ABS(fX2) > DL_FIN_LIM) OR (ABS(fY2) > DL_FIN_LIM) THEN
    bError := TRUE;                 // 量级非有限 / the magnitude is not finite
    RETURN;
END_IF

// 段 3｜对角顶点归一：宽高为负说明录入顺序相反，交换即可 / segment 3, normalise the two corners
fMinX := MIN(fX1, fX2);             // X 下界 / lower X bound
fMaxX := MAX(fX1, fX2);             // X 上界 / upper X bound
fMinY := MIN(fY1, fY2);             // Y 下界 / lower Y bound
fMaxY := MAX(fY1, fY2);             // Y 上界 / upper Y bound
IF ((fMaxX - fMinX) < DL_EPS) AND ((fMaxY - fMinY) < DL_EPS) THEN
    bError := TRUE;                 // 两顶点重合，矩形退化 / the corners coincide and the rectangle degenerates
    RETURN;
END_IF

// 段 4｜四点窗口判定：全走容差窗口，不使用等号 / segment 4, the four sided tolerance window
IF ((fPx > (fMinX - DL_EPS)) AND (fPx < (fMaxX + DL_EPS))) AND ((fPy > (fMinY - DL_EPS)) AND (fPy < (fMaxY + DL_EPS))) THEN
    FC_DL_GeoPointInRectXY := TRUE; // 落在矩形内（含边界） / inside the rectangle, edges included
END_IF
bValid := TRUE;                     // 判定可用 / the verdict is usable
END_FUNCTION

(* ---- FC_DL_GeoPointLineDist.st ---- *)
(*==============================================================================
 * 组件名称 : FC_DL_GeoPointLineDist ｜ 子库 : DL_MathData ｜ v1.0.0 ｜ 2026-11-24
 * 平台     : CODESYS 3.5 / TwinCAT 3 / InoProShop / Machine Expert（纯 IEC，无厂商库）
 * 功能简介 : 点到「无限长直线」的垂直距离。以叉积面积除底边长度实现：
 *            d = |(B−A) × (P−A)| / |B−A|。用于切割头对刀线偏差、视觉边缘距、
 *            机器人轨迹避让安全距离核算。
 * 契约     : 返回距离（≥ 0，同工程单位）；A、B 重合（|AB| < 1.0E-9）时返回 −1.0、
 *            bError := TRUE、bValid := FALSE；任一点含 NaN 或算得非有限值时同样按故障处置。
 * 依赖     : 无 DL_ 内部依赖（R16 自足实现）；Standard.library: ABS / SQRT
 * 错误码   : R297 零码位范式：eErr 恒 0，仅以 bError / bValid 表达
 * 红线自检 : R1 零全局 R2 零%I/%Q R3 纯IEC R4 NaN 自反判据 + 无穷上界 + 退化前拦、
 *            除法前判底边长 ｜ R5 双语注释 R6 N/A（无状态机）R7 N/A（无定时器/沿实例）
 *            R10 无类型转换 R11 全声明行分号 R15 标识符零保留字冲突 R18 N/A（无 bReset）
 * 遗留假设 : 距离为「无限长直线」口径，不是线段距离；需要线段距离的场合须另行裁剪到端点。
 * 修订历史 : 2026-11-24 R79-A 首版（平面几何族 1/8）
 *============================================================================*)
FUNCTION FC_DL_GeoPointLineDist : LREAL
VAR_INPUT
    fPx     : LREAL;    // 被测点 X 坐标 [mm] / X coordinate of the measured point [mm]
    fPy     : LREAL;    // 被测点 Y 坐标 [mm] / Y coordinate of the measured point [mm]
    fAx     : LREAL;    // 直线第一点 X 坐标 [mm] / X coordinate of the first line point [mm]
    fAy     : LREAL;    // 直线第一点 Y 坐标 [mm] / Y coordinate of the first line point [mm]
    fBx     : LREAL;    // 直线第二点 X 坐标 [mm] / X coordinate of the second line point [mm]
    fBy     : LREAL;    // 直线第二点 Y 坐标 [mm] / Y coordinate of the second line point [mm]
END_VAR
VAR_OUTPUT
    eErr    : UDINT;    // 错误码，零码位范式恒 0 / error id, always zero under the zero-code rule
    bError  : BOOL;     // 退化直线或非有限输入为真 / TRUE on a degenerate line or a non finite input
    bValid  : BOOL;     // 结果可用标志 / result usable flag
END_VAR
VAR CONSTANT
    DL_EPS      : LREAL := 1.0E-9;      // 长度容差，底边短于此值即判重合 [mm] / length tolerance for the degenerate test [mm]
    DL_FIN_LIM  : LREAL := 1.0E308;     // 有限性上界，超过按无穷处置 [mm] / finiteness ceiling [mm]
    DL_NEG_ONE  : LREAL := -1.0;        // 退化返回哨兵 / degenerate sentinel
    DL_ZERO_L   : LREAL := 0.0;         // 实数零哨兵 / real zero sentinel
END_VAR
VAR
    fDx     : LREAL;    // 底边 X 分量 B−A [mm] / X component of the base vector [mm]
    fDy     : LREAL;    // 底边 Y 分量 B−A [mm] / Y component of the base vector [mm]
    fLen    : LREAL;    // 底边长度 |B−A| [mm] / base length [mm]
    fCross  : LREAL;    // 叉积绝对值，等于两倍三角形面积 [mm²] / absolute cross product, twice the triangle area [mm²]
END_VAR

// 段 1｜出口预置 / segment 1, preset the exit
FC_DL_GeoPointLineDist := DL_ZERO_L;    // 缺省距离 0 / default distance zero
eErr   := 0;                            // 零码位范式 / zero-code rule
bError := FALSE;                        // 预置无故障 / preset no fault
bValid := FALSE;                        // 计算完成前不认结果 / unusable until the computation ends

// 段 2｜非有限闸：六个坐标任一为 NaN 即拒（x <> x 自反判据） / segment 2, the non finite gate
IF (fPx <> fPx) OR (fPy <> fPy) OR (fAx <> fAx) OR (fAy <> fAy) OR (fBx <> fBx) OR (fBy <> fBy) THEN
    bError := TRUE;                     // 含非数输入 / a not a number input was seen
    FC_DL_GeoPointLineDist := DL_NEG_ONE;
    RETURN;
END_IF

// 段 3｜底边与退化判定：短于容差即两点重合，直线不存在 / segment 3, the base vector and the degenerate test
fDx  := fBx - fAx;                      // X 分量 / the X component
fDy  := fBy - fAy;                      // Y 分量 / the Y component
fLen := SQRT((fDx * fDx) + (fDy * fDy));    // 底边长度，平方和可能溢出为无穷，下一段接住 / the squares may overflow, the next gate catches it
IF (fLen <> fLen) OR (fLen > DL_FIN_LIM) THEN
    bError := TRUE;                     // 长度非有限（坐标量级过大）/ the length is not finite because the coordinates are huge
    FC_DL_GeoPointLineDist := DL_NEG_ONE;
    RETURN;
END_IF
IF fLen < DL_EPS THEN
    bError := TRUE;                     // A、B 重合，直线退化 / the two points coincide and the line degenerates
    FC_DL_GeoPointLineDist := DL_NEG_ONE;
    RETURN;
END_IF

// 段 4｜叉积面积与距离：除法分母已在段 3 证为非零且有限 / segment 4, the cross product and the division
fCross := ABS((fDx * (fPy - fAy)) - (fDy * (fPx - fAx)));   // 两倍三角形面积 / twice the triangle area
IF (fCross <> fCross) OR (fCross > DL_FIN_LIM) THEN
    bError := TRUE;                     // 叉积非有限 / the cross product is not finite
    FC_DL_GeoPointLineDist := DL_NEG_ONE;
    RETURN;
END_IF
FC_DL_GeoPointLineDist := fCross / fLen;    // 面积除底边即高 [mm] / area over base gives the height [mm]
bValid := TRUE;                             // 结果可用 / the result is usable
END_FUNCTION

(* ---- FC_DL_GeoPointRotateXY.st ---- *)
(*==============================================================================
 * 组件名称 : FC_DL_GeoPointRotateXY ｜ 子库 : DL_MathData ｜ v1.0.1 ｜ 2026-11-24
 * 平台     : CODESYS 3.5 / TwinCAT 3 / InoProShop / Machine Expert（纯 IEC，无厂商库）
 * 功能简介 : 平面点绕任意中心旋转。绕 (fCx, fCy) 把点 (fPx, fPy) 逆时针旋转 fAngleDeg 度
 *            （顺时针给负角），输出旋转后坐标。供相机像素坐标与机械坐标对齐、视觉纠偏、
 *            托盘位姿变换使用。
 * 契约     : 入参全有限 → 返回 TRUE、bValid := TRUE、出参有效；任一入参非有限 →
 *            返回 FALSE、bError := TRUE、两出参置 0。角度按 360 取模（负角与超圈角均合法）。
 * 依赖     : 无 DL_ 内部依赖（R16 自足实现），仅用标准库 COS / SIN / TRUNC
 * 错误码   : R297 零码位范式：eErr 恒 0，仅以 bError / bValid 表达
 * 红线自检 : R1 零全局 R2 零%I/%Q R3 纯IEC R4 非有限拦截 + 居中平移后再转（大坐标不丢精度）
 *            R5 双语注释 R6 N/A（无状态机）R7 N/A（无定时器/沿实例）
 *            R10 无类型转换（取整用 TRUNC 泛型）R11 全声明行分号 R15 标识符零保留字冲突
 * 遗留假设 : COS / SIN 取 IEC 61131-3 标准库同名函数（Standard.library），三平台语义一致；
 *            π 内联于常量表，不引用任何度弧换算件；逆时针为正角，与右手坐标系一致，
 *            若目标平台为左手系（Y 向下），调用方取负角即等价。
 * 修订历史 : 2026-11-24 R79-B 首版（几何族 3/3）
 *============================================================================*)
FUNCTION FC_DL_GeoPointRotateXY : BOOL
VAR_INPUT
    fPx       : LREAL := 0.0; // 待旋转点 X 坐标 [mm] / the X coordinate of the point
    fPy       : LREAL := 0.0; // 待旋转点 Y 坐标 [mm] / the Y coordinate of the point
    fAngleDeg : LREAL := 0.0; // 旋转角，逆时针为正，按 360 取模 [度] / the rotation angle, counter clockwise positive, wrapped by 360
    fCx       : LREAL := 0.0; // 旋转中心 X 坐标 [mm] / the X coordinate of the rotation centre
    fCy       : LREAL := 0.0; // 旋转中心 Y 坐标 [mm] / the Y coordinate of the rotation centre
END_VAR
VAR_OUTPUT
    eErr   : UDINT; // 错误码，零码位范式恒 0 / error id, always zero under the zero-code rule
    bError : BOOL;  // 任一入参非有限时为真 / TRUE when any input is not finite
    bValid : BOOL;  // 出参可用标志 / TRUE when the outputs are usable
    fOx    : LREAL; // 旋转后 X 坐标 [mm] / the rotated X coordinate
    fOy    : LREAL; // 旋转后 Y 坐标 [mm] / the rotated Y coordinate
END_VAR
VAR CONSTANT
    DL_FIN     : LREAL := 1.0E30;  // 有限性判据上界（R477 范式：ABS(x)>FIN 判 Inf，禁用 x-x 差判）/ finiteness ceiling, ABS(x)>FIN flags Inf
    DL_ZERO : LREAL := 0.0;               // 实数零哨兵 [mm] / the real zero sentinel
    DL_FULL : LREAL := 360.0;             // 整圆角度 [度] / the full turn in degrees
    DL_DEG  : LREAL := 180.0;             // 半圆角度，度弧换算分母 [度] / the half turn, the divisor of the degree to radian chain
    DL_PI   : LREAL := 3.141592653589793; // 圆周率（内联）[无量纲] / the inline constant pi
END_VAR
VAR
    fTurns : LREAL; // 整圈数（向零截断）[圈] / the whole turn count truncated toward zero
    fAng   : LREAL; // 归一后的旋转角 [度] / the wrapped rotation angle
    fRad   : LREAL; // 旋转角弧度值 [弧度] / the rotation angle in radians
    fCos   : LREAL; // 余弦中间量 [无量纲] / the cosine term
    fSin   : LREAL; // 正弦中间量 [无量纲] / the sine term
    fDx    : LREAL; // 点相对中心的 X 偏移 [mm] / the X offset from the centre
    fDy    : LREAL; // 点相对中心的 Y 偏移 [mm] / the Y offset from the centre
END_VAR

// 段 1｜出口预置 / segment 1, preset the exit
FC_DL_GeoPointRotateXY := FALSE;  // 缺省失败 / default failure
eErr   := 0;                      // 零码位范式 / zero-code rule
bError := FALSE;                  // 预置无故障 / preset no fault
bValid := FALSE;                  // 域闸前不认出参 / the outputs are unusable until the gates pass
fOx    := DL_ZERO;                // X 出参清零 / clear the rotated X
fOy    := DL_ZERO;                // Y 出参清零 / clear the rotated Y

// 段 2｜非有限拦截（五个入参逐个自检，NaN 自反判 + Inf 自减判）/ segment 2, the non finite gate
IF (fPx <> fPx) OR (fPy <> fPy) OR (fAngleDeg <> fAngleDeg) OR (fCx <> fCx) OR (fCy <> fCy) THEN
    bError := TRUE;               // NaN 入参 / a NaN input
    RETURN;                       // 出参保持 0 / the outputs stay zero
END_IF
IF (ABS(fPx) > DL_FIN) OR (ABS(fPy) > DL_FIN) OR (ABS(fAngleDeg) > DL_FIN) OR (ABS(fCx) > DL_FIN) OR (ABS(fCy) > DL_FIN) THEN
    bError := TRUE;               // Inf 入参 / an infinite input
    RETURN;                       // 出参保持 0 / the outputs stay zero
END_IF

// 段 3｜角度归一：θ − TRUNC(θ/360) × 360，负向补一圈到 [0,360) / segment 3, the angle wrap
fTurns := TRUNC(fAngleDeg / DL_FULL);          // 整圈数 [圈] / the whole turn count
fAng   := fAngleDeg - (fTurns * DL_FULL);      // 余角，与输入同号 [度] / the remainder carrying the input sign
IF fAng < DL_ZERO THEN fAng := fAng + DL_FULL; END_IF  // 负向补一圈 / add one turn for negative remainders
fRad := fAng * (DL_PI / DL_DEG);               // 度转弧度 [弧度] / the radian value
fCos := COS(fRad);                             // 余弦 [无量纲] / the cosine term
fSin := SIN(fRad);                             // 正弦 [无量纲] / the sine term

// 段 4｜居中平移后再旋转：先减中心，避免大坐标直接参与乘法丢有效位 / segment 4, the centred rotation
fDx := fPx - fCx;                              // X 偏移 [mm] / the X offset
fDy := fPy - fCy;                              // Y 偏移 [mm] / the Y offset
fOx := fCx + (fDx * fCos) - (fDy * fSin);      // 旋转后 X [mm] / the rotated X
fOy := fCy + (fDx * fSin) + (fDy * fCos);      // 旋转后 Y [mm] / the rotated Y

// 段 5｜出口 / segment 5, the exit
bValid := TRUE;                   // 出参可用 / the outputs are usable
FC_DL_GeoPointRotateXY := TRUE;   // 旋转完成 / the rotation completed
END_FUNCTION

(* ---- FC_DL_GeoPolylineLenFixed.st ---- *)
(*==============================================================================
 * 组件名称 : FC_DL_GeoPolylineLenFixed ｜ 子库 : DL_MathData ｜ v1.0.0 ｜ 2026-11-24
 * 平台     : CODESYS 3.5 / TwinCAT 3 / InoProShop / Machine Expert（纯 IEC，无厂商库）
 * 功能简介 : 定长点列折线总长。两轴坐标以并列定长数组给出，逐段取欧氏距离累加。
 *            用于示教轨迹余量核算、皮带测绘线长、切割路径周长统计。
 * 契约     : 返回折线总长（≥ 0）；nCnt 大于 10 时钳到 10 继续计算（钳位值仍为确定结论，
 *            不置 bError）；nCnt 小于 2 时返回 0 且 bError := TRUE。
 *            数组定长 ARRAY[1..10]，禁变长形参（R17）。
 * 依赖     : 无 DL_ 内部依赖（R16 自足实现）；Standard.library: SQRT
 * 错误码   : R297 零码位范式：eErr 恒 0，仅以 bError / bValid 表达
 * 红线自检 : R1 零全局 R2 零%I/%Q R3 纯IEC R4 点数先钳位后进循环、循环上界由钳位保证
 *            R5 双语注释 R6 N/A（无状态机）R7 N/A（无定时器/沿实例）
 *            R10 无类型转换 R11 全声明行分号 R15 标识符零保留字冲突
 *            R17 定长数组 R18 N/A（无 bReset）
 * 遗留假设 : 数组下标一律从 1 起，与 IEC 默认下界一致；调用方须保证实参数组同为 1..10。
 * 修订历史 : 2026-11-24 R79-A 首版（平面几何族 6/8）
 *============================================================================*)
FUNCTION FC_DL_GeoPolylineLenFixed : LREAL
VAR_INPUT
    aPtsX   : ARRAY[1..10] OF LREAL;    // 点列 X 坐标，1..10 定长 [mm] / X coordinates of the points, fixed length [mm]
    aPtsY   : ARRAY[1..10] OF LREAL;    // 点列 Y 坐标，1..10 定长 [mm] / Y coordinates of the points, fixed length [mm]
    nCnt    : INT;                      // 有效点数，2~10，越界钳位 [个] / effective point count from two to ten, clamped [count]
END_VAR
VAR_OUTPUT
    eErr    : UDINT;    // 错误码，零码位范式恒 0 / error id, always zero under the zero-code rule
    bError  : BOOL;     // 有效点数不足两点为真 / TRUE when fewer than two points remain
    bValid  : BOOL;     // 结果可用标志 / result usable flag
END_VAR
VAR CONSTANT
    DL_PTS_MAX : INT := 10;         // 点列定长上限 [个] / fixed capacity of the point arrays [count]
    DL_PTS_MIN : INT := 2;          // 构成折线的最少点数 [个] / minimum points that form a polyline [count]
    DL_ONE     : INT := 1;          // 下标步长与 1 基起始 [个] / index step and the one based start [count]
    DL_ZERO_L  : LREAL := 0.0;      // 实数零哨兵 [mm] / real zero sentinel [mm]
END_VAR
VAR
    nUse    : INT;      // 钳位后的有效点数 [个] / effective point count after clamping [count]
    i       : INT;      // 段游标，1 起 [个] / segment cursor starting at one [count]
    fDx     : LREAL;    // 单段 X 分量 [mm] / X component of one segment [mm]
    fDy     : LREAL;    // 单段 Y 分量 [mm] / Y component of one segment [mm]
    fSeg    : LREAL;    // 单段长度 [mm] / length of one segment [mm]
    fSum    : LREAL;    // 总长累加器 [mm] / accumulated total length [mm]
END_VAR

// 段 1｜出口预置 / segment 1, preset the exit
FC_DL_GeoPolylineLenFixed := DL_ZERO_L;     // 缺省总长 0 / default total length zero
eErr   := 0;                                // 零码位范式 / zero-code rule
bError := FALSE;                            // 预置无故障 / preset no fault
bValid := FALSE;                            // 计算完成前不认结果 / unusable until the walk ends
fSum   := DL_ZERO_L;                        // 累加器清零 / clear the accumulator

// 段 2｜点数钳位：上越界静默钳位，下越界按故障退出 / segment 2, clamp the point count
nUse := nCnt;                               // 工作副本 / working copy
IF nUse > DL_PTS_MAX THEN
    nUse := DL_PTS_MAX;                     // 钳到定长上限，超出部分不可见 / clamp to the fixed capacity
END_IF
IF nUse < DL_PTS_MIN THEN
    bError := TRUE;                         // 不足两点构不成折线 / fewer than two points form no polyline
    RETURN;                                 // 返回 0 / return zero
END_IF

// 段 3｜逐段累加：下标范围由钳位保证，不会越界 / segment 3, accumulate segment by segment
FOR i := DL_ONE TO (nUse - DL_ONE) DO
    fDx  := aPtsX[i + DL_ONE] - aPtsX[i];                   // X 分量 / X component
    fDy  := aPtsY[i + DL_ONE] - aPtsY[i];                   // Y 分量 / Y component
    fSeg := SQRT((fDx * fDx) + (fDy * fDy));                // 欧氏段长，非有限段由出口自证拦下 / Euclidean length, verified at the exit
    fSum := fSum + fSeg;                                    // 累加 / accumulate
END_FOR

// 段 4｜出口自证：总长必须有限且非负 / segment 4, the exit self proof
IF (fSum <> fSum) OR (fSum < DL_ZERO_L) THEN
    bError := TRUE;                         // 累加结果非有限或为负（坐标量级过大）/ the sum is not finite or negative
    FC_DL_GeoPolylineLenFixed := DL_ZERO_L;
    RETURN;
END_IF
FC_DL_GeoPolylineLenFixed := fSum;          // 总长 / the total length
bValid := TRUE;                             // 结果可用 / the result is usable
END_FUNCTION

(* ---- FC_DL_GrindSpecificEnergyCalc.st ---- *)
(*
  DL Factory R88 | FC_DL_GrindSpecificEnergyCalc
  功能：算比磨削能 u=P/Qw，其中 Qw=ae·vf·b（mm³/s），功率 kW 按 ×1000 换 W，超 60 J/mm³ 提示
  开源溯源：无（clean-room 自研，依据公开工艺公式 比磨削能定义式 u=P/Qw，许可证=MIT，借鉴点=公式结构）
  规则：R1-R16 全遵守；R88 简单件标量形（纯标量入参出参，无循环体、无方法、无属性、无数组）
*)
FUNCTION FC_DL_GrindSpecificEnergyCalc : REAL
VAR_INPUT
    fPowerKW : REAL := 5.0; // 磨削净功率 P（扣除空载） [kW] / net grinding power [kW]
    fAeMm : REAL := 0.02; // 径向切深 ae [mm] / radial depth of cut [mm]
    fVfMmPerS : REAL := 30.0; // 工件进给速度 vf [mm/s] / workpiece feed speed [mm/s]
    fWidthMm : REAL := 20.0; // 磨削接触宽度 b [mm] / grinding contact width [mm]
    fHighLimitJPerMm3 : REAL := 60.0; // 比能偏高阈值（烧伤风险提示） [J/mm³] / high specific energy limit [J/mm^3]
END_VAR
VAR_OUTPUT
    fEnergyJPerMm3 : REAL; // 比磨削能 u [J/mm³] / specific grinding energy [J/mm^3]
    xHigh : BOOL; // TRUE=比能高于阈值，存在烧伤风险 [-] / TRUE when above the limit [-]
END_VAR
VAR
    fPowerW : REAL; // 功率换算为 W [W] / power in watts [W]
    fQwMm3PerS : REAL; // 材料去除率 Qw（除零判据） [mm³/s] / material removal rate, the divisor [mm^3/s]
END_VAR

// 段 1｜出口预置
FC_DL_GrindSpecificEnergyCalc := -1.0; // 哨兵返回 -1（无效） [-] / sentinel return -1, invalid [-]
fEnergyJPerMm3 := 0.0; // 比能预置零 [J/mm³] / specific energy preset zero [J/mm^3]
xHigh := FALSE; // 偏高位预置 FALSE（未判定前不报警） [-] / high flag preset false [-]
fPowerW := 0.0; // 功率 W 值预置零 [W] / power in watts preset zero [W]
fQwMm3PerS := 0.0; // 去除率预置零 [mm³/s] / removal rate preset zero [mm^3/s]

// 段 2｜非有限拦截 + 域闸
IF NOT (fPowerKW > -1.0E30 AND fPowerKW < 1.0E30) OR NOT (fAeMm > -1.0E30 AND fAeMm < 1.0E30) THEN
    RETURN; // 功率/切深任一非有限即拒算 [-] / any non finite input rejected [-]
END_IF
IF NOT (fVfMmPerS > -1.0E30 AND fVfMmPerS < 1.0E30) OR NOT (fWidthMm > -1.0E30 AND fWidthMm < 1.0E30) THEN
    RETURN; // 进给速度/接触宽度任一非有限即拒算 [-] / any non finite input rejected [-]
END_IF
IF NOT (fHighLimitJPerMm3 > -1.0E30 AND fHighLimitJPerMm3 < 1.0E30) THEN
    RETURN; // 阈值非有限则偏高判据失效，故先拦 [J/mm³] / the limit must be finite [J/mm^3]
END_IF
IF fPowerKW < 0.0 OR fAeMm < 0.0 OR fVfMmPerS < 0.0 OR fWidthMm < 1.0E-9 THEN
    RETURN; // 功率/切深/进给非负闸 + 宽度正域闸（分母不得为零） [kW, mm] / non negative terms and positive width
END_IF
IF fHighLimitJPerMm3 <= 0.0 THEN
    RETURN; // 阈值正域闸：非正阈值会使提示恒真 [J/mm³] / positive limit gate [J/mm^3]
END_IF

// 段 3｜计算
fPowerW := fPowerKW * 1000.0; // kW × 1000 W/kW = W，量纲换算 [W] / [kW] x [W/kW] = [W]
fQwMm3PerS := fAeMm * fVfMmPerS * fWidthMm; // mm × (mm/s) × mm = mm³/s，Qw=ae·vf·b / [mm^3/s]
IF fQwMm3PerS < 1.0E-9 THEN
    RETURN; // 除法前分母闸：去除率须大于 1E-9（零切深会除零） [mm³/s] / denominator gate [mm^3/s]
END_IF
fEnergyJPerMm3 := fPowerW / fQwMm3PerS; // (J/s) ÷ (mm³/s) = J/mm³，即比磨削能 [J/mm³] / [J/mm^3]

// 段 4｜判定与饱和
IF NOT (fEnergyJPerMm3 > -1.0E30 AND fEnergyJPerMm3 < 1.0E30) THEN
    RETURN; // 结果非有限再拦一次 [-] / re-check the result for finiteness [-]
END_IF
xHigh := fEnergyJPerMm3 > fHighLimitJPerMm3; // 严格大于阈值为偏高，等于阈值仍判正常 [J/mm³] / strict compare [J/mm^3]

// 段 5｜出口自检
IF fEnergyJPerMm3 < 0.0 THEN
    RETURN; // 出口自检：比能不得为负（负值说明功率符号错） [J/mm³] / energy must not be negative [J/mm^3]
END_IF
FC_DL_GrindSpecificEnergyCalc := fEnergyJPerMm3; // 返回比磨削能 [J/mm³] / return the specific energy [J/mm^3]
END_FUNCTION

(* ---- FC_DL_GrindWheelPeripheralSpeedCalc.st ---- *)
(*
  DL Factory R88 | FC_DL_GrindWheelPeripheralSpeedCalc
  功能：由砂轮直径与转速算外周线速度 v=π·D·n/60000（mm,rpm→m/s），超 35 m/s 报警
  开源溯源：无（clean-room 自研，依据公开工艺公式 砂轮线速度式 v=π·D·n，许可证=MIT，借鉴点=公式结构）
  规则：R1-R16 全遵守；R88 简单件标量形（纯标量入参出参，无循环体、无方法、无属性、无数组）
*)
FUNCTION FC_DL_GrindWheelPeripheralSpeedCalc : REAL
VAR_INPUT
    fDiaMm : REAL := 400.0; // 砂轮外径 D [mm] / wheel outer diameter [mm]
    fRpm : REAL := 1500.0; // 主轴转速 n [r/min] / spindle speed [rpm]
    fLimitMPerS : REAL := 35.0; // 线速度报警阈值（常规树脂结合剂 35 m/s） [m/s] / overspeed alarm limit [m/s]
END_VAR
VAR_OUTPUT
    fSpeedMPerS : REAL; // 砂轮外周线速度 v [m/s] / peripheral speed [m/s]
    xOverLimit : BOOL; // TRUE=线速度超过阈值，需报警 [-] / TRUE when above the alarm limit [-]
END_VAR
VAR
    fCircMMm : REAL; // 单转行程 π·D [mm/rev] / travel per revolution [mm/rev]
    fMMPerMin : REAL; // 每分钟行程 π·D·n [mm/min] / travel per minute [mm/min]
END_VAR

// 段 1｜出口预置
FC_DL_GrindWheelPeripheralSpeedCalc := -1.0; // 哨兵返回 -1（无效） [-] / sentinel return -1, invalid [-]
fSpeedMPerS := 0.0; // 线速度预置零 [m/s] / speed preset zero [m/s]
xOverLimit := FALSE; // 超限位预置 FALSE（未判定前不报超限） [-] / over-speed flag preset false [-]
fCircMMm := 0.0; // 单转行程预置零 [mm/rev] / circumference preset zero [mm/rev]
fMMPerMin := 0.0; // 每分钟行程预置零 [mm/min] / travel per minute preset zero [mm/min]

// 段 2｜非有限拦截 + 域闸
IF NOT (fDiaMm > -1.0E30 AND fDiaMm < 1.0E30) OR NOT (fRpm > -1.0E30 AND fRpm < 1.0E30) THEN
    RETURN; // 直径/转速任一非有限即拒算 [-] / any non finite input rejected [-]
END_IF
IF NOT (fLimitMPerS > -1.0E30 AND fLimitMPerS < 1.0E30) THEN
    RETURN; // 阈值非有限则报警判据失效，故先拦 [m/s] / the alarm limit must be finite [m/s]
END_IF
IF fDiaMm < 1.0E-9 OR fRpm < 0.0 THEN
    RETURN; // 直径正域闸 + 转速非负闸 [mm, r/min] / positive diameter and non negative speed
END_IF
IF fLimitMPerS <= 0.0 THEN
    RETURN; // 阈值正域闸：非正阈值会使报警恒真或恒假 [m/s] / positive limit gate [m/s]
END_IF

// 段 3｜计算
fCircMMm := 3.14159265 * fDiaMm; // 无量纲 × mm = mm/rev，每转行程 π·D [mm/rev] / [mm] per revolution
fMMPerMin := fCircMMm * fRpm; // (mm/rev) × (r/min) = mm/min，每分钟行程 [mm/min] / [mm/min]
fSpeedMPerS := fMMPerMin / 60000.0; // (mm/min) ÷ 60000 = m/s；60000=1000 mm/m × 60 s/min 恒正 [m/s] / [m/s]

// 段 4｜判定与饱和
IF NOT (fSpeedMPerS > -1.0E30 AND fSpeedMPerS < 1.0E30) THEN
    RETURN; // 结果非有限再拦一次（防溢出成 Inf） [m/s] / re-check the result for finiteness [m/s]
END_IF
xOverLimit := fSpeedMPerS > fLimitMPerS; // 严格大于阈值为超限，等于阈值仍判合格 [m/s] / strict compare against the limit [m/s]

// 段 5｜出口自检
IF fSpeedMPerS < 0.0 THEN
    RETURN; // 出口自检：线速度不得为负（负值说明输入符号错） [m/s] / speed must not be negative [m/s]
END_IF
FC_DL_GrindWheelPeripheralSpeedCalc := fSpeedMPerS; // 返回砂轮线速度 [m/s] / return the peripheral speed [m/s]
END_FUNCTION

(* ---- FC_DL_H2LeakRateCalc.st ---- *)
(*
  DL Factory R88 | FC_DL_H2LeakRateCalc
  功能：压降法算泄漏率 Q=V·Δp/Δt（Pa·m³/s），换算为标准状态 NmL/min，并判是否超限
  开源溯源：无（clean-room 自研，依据公开工艺公式 压降法泄漏率式 Q=V·dp/dt，许可证=MIT，借鉴点=公式结构）
  规则：R1-R16 全遵守；R88 简单件标量形（纯标量入参出参，无循环体、无方法、无属性、无数组）
*)
FUNCTION FC_DL_H2LeakRateCalc : REAL
VAR_INPUT
    fVolL : REAL := 50.0; // 被测封闭容积 V [L] / test volume [L]
    fDropPa : REAL := 500.0; // 保压期间压降 Δp（取正值） [Pa] / pressure drop over the hold time [Pa]
    fDurS : REAL := 60.0; // 保压时长 Δt [s] / hold duration [s]
    fLimitNmlMin : REAL := 10.0; // 泄漏率报警上限（标准状态） [NmL/min] / leak rate alarm limit [NmL/min]
    fPatmPa : REAL := 101325.0; // 标准大气压（换算基准） [Pa] / standard atmospheric pressure [Pa]
END_VAR
VAR_OUTPUT
    fLeakNmlMin : REAL; // 泄漏率（标准状态体积流量） [NmL/min] / leak rate at standard conditions [NmL/min]
    xOverLimit : BOOL; // TRUE=泄漏率超过报警上限 [-] / TRUE when above the alarm limit [-]
END_VAR
VAR
    fVolM3 : REAL; // 容积换算为 m³ [m³] / volume in cubic metres [m^3]
    fLeakPam3PerS : REAL; // 泄漏率原始量 Q [Pa·m³/s] / raw leak rate [Pa*m^3/s]
    fLeakNm3PerS : REAL; // 标准状态体积流量 [Nm³/s] / standard volumetric flow [Nm^3/s]
END_VAR

// 段 1｜出口预置
FC_DL_H2LeakRateCalc := -1.0; // 哨兵返回 -1（无效） [-] / sentinel return -1, invalid [-]
fLeakNmlMin := 0.0; // 泄漏率预置零 [NmL/min] / leak rate preset zero [NmL/min]
xOverLimit := FALSE; // 超限位预置 FALSE（未判定前不报警） [-] / over-limit flag preset false [-]

// 段 2｜非有限拦截 + 域闸
IF NOT (fVolL > -1.0E30 AND fVolL < 1.0E30) OR NOT (fDropPa > -1.0E30 AND fDropPa < 1.0E30) OR NOT (fDurS > -1.0E30 AND fDurS < 1.0E30) THEN
    RETURN; // 容积/压降/时长任一非有限即拒算 [-] / any non finite input rejected [-]
END_IF
IF NOT (fLimitNmlMin > -1.0E30 AND fLimitNmlMin < 1.0E30) OR NOT (fPatmPa > -1.0E30 AND fPatmPa < 1.0E30) THEN
    RETURN; // 上限/基准压力任一非有限则判据与换算链失效，故先拦 [-] / these pins must be finite [-]
END_IF
IF fVolL < 1.0E-9 OR fDropPa < 0.0 OR fDurS < 1.0E-9 THEN
    RETURN; // 容积正域闸 + 压降非负闸 + 时长正域闸（分母不得为零） [L, Pa, s] / positive volume and duration
END_IF
IF fPatmPa < 1.0E-9 OR fLimitNmlMin <= 0.0 THEN
    RETURN; // 基准压力正域闸（换算分母）+ 上限正域闸 [Pa, NmL/min] / reference pressure and limit gates
END_IF

// 段 3｜计算（Pa·m³/s → Nm³/s → NmL/min 三段换算，逐项量纲见行尾注释）
fVolM3 := fVolL * 0.001; // L × 0.001 m³/L = m³，容积换算 [m³] / [L] x [m^3/L] = [m^3]
fLeakPam3PerS := fVolM3 * fDropPa / fDurS; // m³ × Pa ÷ s = Pa·m³/s，压降法泄漏率 [Pa·m³/s] / [Pa*m^3/s]
fLeakNm3PerS := fLeakPam3PerS / fPatmPa; // (Pa·m³/s) ÷ Pa = m³/s（标准状态） [Nm³/s] / [Nm^3/s]
fLeakNmlMin := fLeakNm3PerS * 1.0E6 * 60.0; // (Nm³/s) × 1e6 mL/m³ × 60 s/min = NmL/min [NmL/min] / [NmL/min]

// 段 4｜判定与饱和
IF NOT (fLeakNmlMin > -1.0E30 AND fLeakNmlMin < 1.0E30) THEN
    RETURN; // 结果非有限再拦一次 [-] / re-check the result for finiteness [-]
END_IF
xOverLimit := fLeakNmlMin > fLimitNmlMin; // 严格大于上限为超限，等于上限仍判合格 [NmL/min] / strict compare [NmL/min]

// 段 5｜出口自检
IF fLeakNmlMin < 0.0 THEN
    RETURN; // 出口自检：泄漏率不得为负（负值说明压降符号错） [NmL/min] / leak rate must not be negative [NmL/min]
END_IF
FC_DL_H2LeakRateCalc := fLeakNmlMin; // 返回标准状态泄漏率 [NmL/min] / return the leak rate [NmL/min]
END_FUNCTION

(* ---- FC_DL_HaversineDistance.st ---- *)
(*
  Name        : FC_DL_HaversineDistance
  Category    : DL_MathData
  Version     : 1.0.0
  Purpose     : 球面两点大圆距离（Haversine 公式，双精度），供 AGV/巡检定位换算；输入为十进制度，输出为米；/ Great-circle distance between two points via the Haversine formula in double precision; inputs in decimal degrees, output in metres
  溯源        : t2-1-lgf-math ◐/自研，clean-room 实现
  Boundary    : ① 入口有限性闸：任一输入 NaN（x = x 自反）或 Inf（(x-x) = (x-x) 差判）→ bValid = FALSE，返回 0.0（哨兵零点）；
                ② 输入域钳位：纬度钳 -90..90，经度差归一化到 -180..180（不钳位经度本身，跨 180° 子午线正确）；
                ③ 除零前置：公式内除子为常量（2/半径换算）与 asin 域保护（根号项钳 0..1）；
                ④ 钳位是各中间量的最后一次写（纬度/经度差/根号项），钳完不被覆盖；
                ⑤ 返回值 = 两点球面距离 [m]，bValid = FALSE 时不得使用返回值（上层契约）。
*)
FUNCTION FC_DL_HaversineDistance : LREAL
VAR_INPUT
    fLat1 : LREAL;                           (* 点 1 纬度，域 -90..90（越域钳位）[°] / Point 1 latitude *)
    fLon1 : LREAL;                           (* 点 1 经度 [°] / Point 1 longitude *)
    fLat2 : LREAL;                           (* 点 2 纬度，域 -90..90（越域钳位）[°] / Point 2 latitude *)
    fLon2 : LREAL;                           (* 点 2 经度 [°] / Point 2 longitude *)
END_VAR
VAR_OUTPUT
    bValid : BOOL;                           (* 结果有效标志（FALSE 时返回值为哨兵零点）[-] / Result validity flag *)
END_VAR
VAR CONSTANT
    DL_HAV_R_EARTH : LREAL := 6371008.8;     (* 地球平均半径 [m] / Earth mean radius *)
    DL_HAV_DEG2RAD : LREAL := 0.017453292519943295;   (* 度→弧度换算常量 π/180 [-] / Degrees to radians factor *)
    DL_HAV_LATMAX  : LREAL := 90.0;          (* 纬度钳位绝对值上限 [°] / Latitude clamp magnitude *)
    DL_HAV_LONSPAN : LREAL := 360.0;         (* 经度整圆跨度（归一化用）[°] / Longitude full circle span *)
    DL_HAV_HALF    : LREAL := 0.5;           (* 半角换算常量 [-] / Half factor *)
    DL_HAV_TWO     : LREAL := 2.0;           (* 反正弦倍率常量 [-] / Arc-sine multiplier *)
END_VAR
VAR
    _fLat1   : LREAL;                        (* 钳位后点 1 纬度 [°] / Clamped latitude 1 *)
    _fLat2   : LREAL;                        (* 钳位后点 2 纬度 [°] / Clamped latitude 2 *)
    _fDLon   : LREAL;                        (* 归一化后经度差 [°] / Normalised longitude delta *)
    _fPhi1   : LREAL;                        (* 点 1 纬度弧度 [rad] / Latitude 1 in radians *)
    _fPhi2   : LREAL;                        (* 点 2 纬度弧度 [rad] / Latitude 2 in radians *)
    _fDPhi   : LREAL;                        (* 纬度差弧度 [rad] / Latitude delta radians *)
    _fDLam   : LREAL;                        (* 经度差弧度 [rad] / Longitude delta radians *)
    _fSinDp  : LREAL;                        (* sin(Δφ/2) 中间量 [-] / Half-chord sine term 1 *)
    _fSinDl  : LREAL;                        (* sin(Δλ/2) 中间量 [-] / Half-chord sine term 2 *)
    _fA      : LREAL;                        (* Haversine a 中间量 [-] / Haversine a term *)
    _fC      : LREAL;                        (* Haversine c 中间量（asin 域已钳）[-] / Haversine c term *)
END_VAR

(* —— 段 0：入口有限性闸（NaN 自反 + Inf 差判，四输入逐项） —— *)
bValid := TRUE;                                                                (* 有效标志预置（任一闸命中即翻 FALSE） / Validity preset *)
IF NOT ((fLat1 = fLat1) AND ((fLat1 - fLat1) = (fLat1 - fLat1))) THEN
    bValid := FALSE;                                                           (* 纬度 1 非有限 / Latitude 1 non-finite *)
END_IF
IF NOT ((fLon1 = fLon1) AND ((fLon1 - fLon1) = (fLon1 - fLon1))) THEN
    bValid := FALSE;                                                           (* 经度 1 非有限 / Longitude 1 non-finite *)
END_IF
IF NOT ((fLat2 = fLat2) AND ((fLat2 - fLat2) = (fLat2 - fLat2))) THEN
    bValid := FALSE;                                                           (* 纬度 2 非有限 / Latitude 2 non-finite *)
END_IF
IF NOT ((fLon2 = fLon2) AND ((fLon2 - fLon2) = (fLon2 - fLon2))) THEN
    bValid := FALSE;                                                           (* 经度 2 非有限 / Longitude 2 non-finite *)
END_IF

(* —— 段 1：无效输入早退（返回哨兵零点） —— *)
IF NOT bValid THEN
    FC_DL_HaversineDistance := 0.0;                                            (* 哨兵零点返回 / Sentinel zero return *)
    RETURN;
END_IF

(* —— 段 2：输入域钳位与经度差归一化（各自中间量最后一次写） —— *)
_fLat1 := fLat1;                                                               (* 点 1 纬度装载 / Load latitude 1 *)
IF _fLat1 > DL_HAV_LATMAX THEN
    _fLat1 := DL_HAV_LATMAX;                                                   (* 纬度上限钳位 / Latitude upper clamp *)
END_IF
IF _fLat1 < -DL_HAV_LATMAX THEN
    _fLat1 := -DL_HAV_LATMAX;                                                  (* 纬度下限钳位 / Latitude lower clamp *)
END_IF
_fLat2 := fLat2;                                                               (* 点 2 纬度装载 / Load latitude 2 *)
IF _fLat2 > DL_HAV_LATMAX THEN
    _fLat2 := DL_HAV_LATMAX;                                                   (* 纬度上限钳位 / Latitude upper clamp *)
END_IF
IF _fLat2 < -DL_HAV_LATMAX THEN
    _fLat2 := -DL_HAV_LATMAX;                                                  (* 纬度下限钳位 / Latitude lower clamp *)
END_IF
_fDLon := fLon2 - fLon1;                                                       (* 原始经度差 [°] / Raw longitude delta *)
_fDLon := _fDLon - DL_HAV_LONSPAN * TRUNC(_fDLon / DL_HAV_LONSPAN);            (* 整圈折返到 (-360, 360)（除子为常量） / Fold into one circle *)
IF _fDLon > 180.0 THEN
    _fDLon := _fDLon - DL_HAV_LONSPAN;                                         (* 折回 (-180, 180]，跨 180° 子午线正确 / Fold back across antimeridian *)
ELSIF _fDLon <= -180.0 THEN
    _fDLon := _fDLon + DL_HAV_LONSPAN;                                         (* 折回 (-180, 180] / Fold back *)
END_IF

(* —— 段 3：Haversine 公式本体（除子全为常量，无运行期除零） —— *)
_fPhi1 := _fLat1 * DL_HAV_DEG2RAD;                                             (* 点 1 纬度弧度 [rad] / Latitude 1 radians *)
_fPhi2 := _fLat2 * DL_HAV_DEG2RAD;                                             (* 点 2 纬度弧度 [rad] / Latitude 2 radians *)
_fDPhi := (_fLat2 - _fLat1) * DL_HAV_DEG2RAD;                                  (* 纬度差弧度 [rad] / Latitude delta radians *)
_fDLam := _fDLon * DL_HAV_DEG2RAD;                                             (* 经度差弧度 [rad] / Longitude delta radians *)
_fSinDp := SIN(_fDPhi * DL_HAV_HALF);                                          (* sin(Δφ/2) [-] / Sine term 1 *)
_fSinDl := SIN(_fDLam * DL_HAV_HALF);                                          (* sin(Δλ/2) [-] / Sine term 2 *)
_fA := _fSinDp * _fSinDp + COS(_fPhi1) * COS(_fPhi2) * _fSinDl * _fSinDl;      (* Haversine a [-] / Haversine a *)
IF _fA > 1.0 THEN
    _fA := 1.0;                                                                (* a 上界钳 1（浮点溢出防护，asin 定义域） / Clamp a to domain *)
ELSIF _fA < 0.0 THEN
    _fA := 0.0;                                                                (* a 下界钳 0（asin 定义域） / Clamp a to domain *)
END_IF
_fC := ASIN(SQRT(_fA)) * DL_HAV_TWO;                                           (* 大圆角距 c（定义域已钳）[rad] / Central angle *)
FC_DL_HaversineDistance := DL_HAV_R_EARTH * _fC;                               (* 球面距离 = R × c [m] / Distance = R times c *)
END_FUNCTION

(* ---- FC_DL_HermiteInterp.st ---- *)
(*
  ==================================================================
  组件名 Component  : FC_DL_HermiteInterp
  分类   Category   : DL_MathData
  复杂度 Complexity  : cx3
  版本   Version    : 1.0.0
  功能   Purpose    : 单区间三次 Hermite 插值。由端点值 y0 / y1 与端点斜率 m0 / m1
                      四条件唯一确定区间 [x0, x1] 内的三次多项式，输出插值 y；
                      x 越出区间按端点钳位并置 bClamped，x1 = x0（含反向）判退化
                      （bDegenerate，出口取 y0），任一输入非有限置 bInvalid 且出口取零。
  来源   Source     : t2-1-lgf-math
  溯源   Origin     : IEC 61131-3 标准语义的道莅防御性实现；三次 Hermite 基函数为公开
                      数值分析结果，clean-room 自研实现，未复制任何闭源代码行。
  平台   Platform   : 纯 IEC 61131-3（LREAL 运算，无私有库、无方言转换、无幂运算符）
  作者   Author     : 道莅代码库 · PLC 编程专家（R56）
  ------------------------------------------------------------------
  边界 Boundary     :
                      一 本件只做单区间插值，不建全局网格表、不做样条全局连续性（属主边界）；
                      二 区间方向固定 x0 < x1，区间宽度不大于 1.0E-12 一律判退化并取 y0；
                      三 非有限输入不穿透出口，安全侧取常量零（R127）；
                      四 早退分支出口变换与主体一致（R94）：退化分支取 y0 即四条件曲线
                         在退化极限下的正确极限值；
                      五 无全局变量、无外部变量声明、无物理地址寻址、无定时器（纯函数）。
  输出契约 Output contract:
                      y 仅在输入有限时为插值结果；标志优先级 bInvalid > bDegenerate > bClamped；
                      本件为纯函数，无跨扫描周期状态驻留。
  修订记录 Revision  :
    2026-11-20  v1.0.0  R56 首版（批 1 · 序号 1）
  ==================================================================
*)

FUNCTION FC_DL_HermiteInterp : LREAL
VAR_INPUT
    x  : LREAL; // 插值自变量 [自变量单位] / independent variable of the interpolation
    x0 : LREAL; // 区间左端点 [自变量单位] / left interval bound
    x1 : LREAL; // 区间右端点 [自变量单位] / right interval bound
    y0 : LREAL; // 左端点函数值 [因变量单位] / function value at the left bound
    y1 : LREAL; // 右端点函数值 [因变量单位] / function value at the right bound
    m0 : LREAL; // 左端点斜率 [因变量每自变量] / slope at the left bound
    m1 : LREAL; // 右端点斜率 [因变量每自变量] / slope at the right bound
END_VAR
VAR_OUTPUT
    bClamped    : BOOL; // x 越出区间已按端点钳位 [-] / x was clamped to an interval bound
    bDegenerate : BOOL; // 区间退化（x1 = x0），出口取 y0 [-] / degenerate interval, the outlet takes y0
    bInvalid    : BOOL; // 任一输入非有限，出口取零 [-] / any input non finite, the outlet takes zero
END_VAR
VAR
    _bFin  : BOOL := FALSE; // 七个输入全部有限 [-] / all seven inputs are finite
    _fDx   : LREAL := 0.0;  // 区间宽度 [自变量单位] / interval width
    _fXUse : LREAL := 0.0;  // 钳位后的插值自变量 [自变量单位] / clamped independent variable
    _fT    : LREAL := 0.0;  // 归一化区间参数（0..1）[无量纲] / normalised interval parameter
    _fT2   : LREAL := 0.0;  // 参数平方 [无量纲] / square of the parameter
    _fT3   : LREAL := 0.0;  // 参数立方 [无量纲] / cube of the parameter
    _fH00  : LREAL := 0.0;  // Hermite 基函数 h00 [无量纲] / Hermite basis h00
    _fH10  : LREAL := 0.0;  // Hermite 基函数 h10 [无量纲] / Hermite basis h10
    _fH01  : LREAL := 0.0;  // Hermite 基函数 h01 [无量纲] / Hermite basis h01
    _fH11  : LREAL := 0.0;  // Hermite 基函数 h11 [无量纲] / Hermite basis h11
END_VAR

// 段 1｜非有限闸（R151 全覆盖）：七个输入逐项判，NaN 自反、Inf 差值自减 / segment 1, finiteness gate over every input
_bFin := (x = x) AND ((x - x) = (x - x)) AND (x0 = x0) AND ((x0 - x0) = (x0 - x0)) AND (x1 = x1) AND ((x1 - x1) = (x1 - x1)) AND (y0 = y0) AND ((y0 - y0) = (y0 - y0)) AND (y1 = y1) AND ((y1 - y1) = (y1 - y1)) AND (m0 = m0) AND ((m0 - m0) = (m0 - m0)) AND (m1 = m1) AND ((m1 - m1) = (m1 - m1)); // 七输入有限性判定 / finiteness verdict over all seven inputs
IF NOT _bFin THEN // 非有限输入 / non finite input
    FC_DL_HermiteInterp := 0.0; // 安全侧取常量零（R127）/ the safe side takes the constant zero
    bInvalid := TRUE; // 置无效标志 / raise the invalid flag
    bClamped := FALSE; // 钳位标志不成立 / the clamp flag is false
    bDegenerate := FALSE; // 退化标志不成立 / the degenerate flag is false
    RETURN; // 早退 / early return
END_IF
bInvalid := FALSE; // 有限输入，无效标志不成立 / finite input, the invalid flag is false

// 段 2｜退化判据：区间宽度不大于退化阈即取左端点值 / segment 2, degeneracy verdict
_fDx := x1 - x0; // 区间宽度 / interval width
IF _fDx <= 1.0E-12 THEN // 区间退化（含反向区间与等端点）/ the interval is degenerate
    FC_DL_HermiteInterp := y0; // 出口取左端点值（四条件曲线的退化极限，R94 一致出口）/ the outlet takes the left bound value, the degenerate limit of the same curve
    bDegenerate := TRUE; // 置退化标志 / raise the degenerate flag
    bClamped := FALSE; // 钳位标志不成立 / the clamp flag is false
    RETURN; // 早退 / early return
END_IF

// 段 3｜越域钳位 / segment 3, domain clamp
_fXUse := x; // 自变量直通 / the abscissa passes through
bClamped := FALSE; // 钳位标志预置假 / preset the clamp flag to false
IF x < x0 THEN // 左越域 / below the left bound
    _fXUse := x0; // 钳到左端点 / clamp to the left bound
    bClamped := TRUE; // 置钳位标志 / raise the clamp flag
ELSIF x > x1 THEN // 右越域 / above the right bound
    _fXUse := x1; // 钳到右端点 / clamp to the right bound
    bClamped := TRUE; // 置钳位标志 / raise the clamp flag
END_IF

// 段 4｜Hermite 基函数与四条件插值（幂次以显式乘法展开，禁 **）/ segment 4, Hermite basis and interpolation with explicit multiplications
_fT := (_fXUse - x0) / _fDx; // 归一化参数，除子为区间宽度已证大于退化阈 / normalised parameter, the divisor is the proven width
_fT2 := _fT * _fT; // 参数平方 / square of the parameter
_fT3 := _fT2 * _fT; // 参数立方 / cube of the parameter
_fH00 := 2.0 * _fT3 - 3.0 * _fT2 + 1.0; // 基函数 h00（端点值权重）/ basis h00, the endpoint value weight
_fH10 := _fT3 - 2.0 * _fT2 + _fT; // 基函数 h10（端点斜率权重）/ basis h10, the endpoint slope weight
_fH01 := -2.0 * _fT3 + 3.0 * _fT2; // 基函数 h01 / basis h01
_fH11 := _fT3 - _fT2; // 基函数 h11 / basis h11
FC_DL_HermiteInterp := _fH00 * y0 + _fH10 * _fDx * m0 + _fH01 * y1 + _fH11 * _fDx * m1; // 四条件三次插值 / the cubic interpolation from four conditions
END_FUNCTION

(* ---- FC_DL_HexStringToBytes.st ---- *)
(*==============================================================================
 * 组件名称 (Component)  : FC_DL_HexStringToBytes
 * 所属子库 (Sublibrary) : DL_MathData
 * 当前版本 (Version)    : 1.0.0
 * 兼容性   (Platform)   : CODESYS 3.5 / TwinCAT 3 / 汇川 InoProShop / Machine Expert
 *                         仅依赖 Standard.library（LEN / MID / FIND / SHL / 显式转换），
 *                         无厂商方言，字符访问用标准 MID 函数而非下标方言
 * 功能描述 (Function)   : 十六进制 ASCII 字符串到字节数组的严格解析。
 *                         "1A2B3C" → 16#1A, 16#2B, 16#3C；可选剥离 Modbus ASCII
 *                         帧的冒号帧头与回车换行帧尾。用于扫码枪十六进制输出、
 *                         Modbus ASCII 收帧、RFID 标签 ID 解析、固件分段校验的
 *                         前置解码。与 FC_DL_LrcChecksum 组成"先解码、后校验"
 *                         的两步收帧链路。
 *                         两遍扫描严格模式：第一遍全量校验字符合法性，
 *                         第二遍才写入输出——任何失败路径不留下半截缓冲。
 *
 * 【严格模式声明 / Strict-mode statement（边界 B2）】
 *   **不跳过空格、不跳过 0x 前缀、不容忍内嵌分隔符**："1A 2B" 判非法。
 *   宽容解析会把组帧错误吃进数据层，现场表现为"校验通过但数据错"，
 *   比直接报错难查一个数量级。
 *
 * 【先校验后写入 / Validate-then-write（边界 B1）】
 *   任何失败路径不得留下部分写入的输出缓冲——调用方可能直接把缓冲
 *   拿去发报文，半截字节流比没有更危险。
 *
 * 【奇数长度 / Odd length（边界 B4）】
 *   判非法而非"末尾补 0"——补 0 会凭空造出一个字节。
 *
 * 【位置语义 / Position semantics（边界 B9）】
 *   nInvalidPos 为原文 1 起的字符位置（含被剥离的冒号），便于现场
 *   拿着报文直接数到出错字符。
 *
 * 【字符串长度警示 / String-length warning（边界 B6）】
 *   形参显式声明为 255 长度：CODESYS 系平台默认 STRING 仅 80 字节，
 *   不显式声明长度会被静默截断，长报文解析出错且无任何提示。
 *
 * 【验收向量 / Acceptance vectors】
 *   V1  "1A2B3C"，nMaxBytes = 64 → 返回 3；[16#1A, 16#2B, 16#3C]
 *   V2  "1a2b"（小写）→ 返回 2；[16#1A, 16#2B]
 *   V3  ":010300000001FB" + CR + LF，bStripFraming = TRUE
 *       → 返回 7；[01,03,00,00,00,01,FB]（与 FC_DL_LrcChecksum V1 闭环）
 *   V4  "1A2B3"（奇数长度）→ 返回 -1、16#0002_000A、nInvalidPos = 6、缓冲不变
 *   V5  "1G"（非法字符）→ 返回 -1、16#0002_000A、nInvalidPos = 2
 *   V6  130 字符（65 字节）且 nMaxBytes = 64 → 返回 -1、16#0001_0009、缓冲不变
 *   V7  空串 → 返回 0、uErrorId = 0（空报文合法，由上层判长度）
 * 开源溯源 (Origin)     : 原创实现（参考西门子 LGF 转换器组"字符串与数值互转、
 *                         按类型分函数、单一职责"的组织方式，以及 Modbus 应用
 *                         协议规范的 ASCII 帧定义，clean-room 编写，
 *                         未复制任何源码）。
 * 依赖     (Depends)    : 无 DL_ 内部依赖（配套校验见 FC_DL_LrcChecksum）
 * 红线自检 (Redline)    : R1 ✓ 零全局变量表与外部变量引用 ｜ R2 ✓ 零物理 IO 地址直写
 *                         R3 ✓ 纯 IEC 61131-3（MID/FIND 取字符，无下标方言、无指针）
 *                         R4 ✓ 容量钳位 + 奇数与非法字符拒绝 + 失败不写缓冲
 *                         R5 ✓ 全变量中英双语同行注释 ｜ R6 N/A（无状态机）｜ R7 N/A（无实例调用）
 * 修订历史 (Revision)   :
 *   2026-11-14  v1.0.0  首版入库（Phase 1 收口批次 · R3）
 *============================================================================*)
FUNCTION FC_DL_HexStringToBytes : INT
VAR_IN_OUT
    aabyOut       : ARRAY[0..63] OF BYTE;   // 输出字节缓冲，失败时不写入 / Output buffer, untouched on failure
END_VAR
VAR_INPUT
    sHex          : STRING(255);            // 十六进制字符串，显式 255 长度防截断 / Hex string, explicit 255 length
    bStripFraming : BOOL := FALSE;          // TRUE：剥离首冒号与尾部回车换行 / TRUE: strip leading colon and trailing CR/LF
    nMaxBytes     : INT  := 64;             // 允许写入的最大字节数，1..64 / Maximum bytes to write, range 1..64
END_VAR
VAR_OUTPUT
    nInvalidPos   : INT;                    // 首个非法字符位置（原文 1 起），0 = 无 / First invalid char position, 1-based in the original
    uErrorId      : UDINT;                  // 故障码，0 = 无故障 / Error code, 0 = no error
END_VAR
VAR
    nLen          : INT;                    // 原文长度 / Original string length
    nStart        : INT;                    // 有效起始位置（1 起） / Effective start index, 1-based
    nEnd          : INT;                    // 有效结束位置（1 起，含） / Effective end index, 1-based inclusive
    nHexLen       : INT;                    // 有效十六进制字符数 / Effective hex character count
    nBytes        : INT;                    // 待写字节数 / Bytes to write
    nI            : INT;                    // 字符或字节循环索引 / Char or byte loop index
    nHiNib        : INT;                    // 高半字节值 0..15 / High nibble value 0..15
    nLoNib        : INT;                    // 低半字节值 0..15 / Low nibble value 0..15
    sChar         : STRING(1);              // 当前字符（标准 MID 取出） / Current char via standard MID
END_VAR
VAR CONSTANT
    DL_HX_BUF_MAX  : INT := 64;             // 输出缓冲上限，必须与数组维度一致 / Output buffer limit, must match the array
    DL_HX_PAIR     : INT := 2;              // 每字节字符数 / Chars per byte
    DL_HX_ONE      : INT := 1;              // MID 单字符长度参数 / MID single-char length
    DL_HX_SHIFT    : INT := 4;              // 高半字节左移位数 / High-nibble shift count
    DL_HX_COLON    : STRING(1) := ':';      // Modbus ASCII 帧头 / Modbus ASCII frame start
    DL_HX_CR       : STRING(1) := '$R';     // 回车 / Carriage return
    DL_HX_LF       : STRING(1) := '$L';     // 换行 / Line feed
    DL_HX_DIG_UP   : STRING := '0123456789ABCDEF'; // 大写十六进制字符表（FIND 定位） / Uppercase hex digits for FIND lookup
    DL_HX_DIG_LOW  : STRING := '0123456789abcdef'; // 小写十六进制字符表（FIND 定位） / Lowercase hex digits for FIND lookup
END_VAR

(*------------------------------------------------------------------------------
 * 段 1｜安全预置：返回值与位置码归零，先校验后写入（边界 B1）
 *      Safe preset: return and position cleared, validate before writing
 *-----------------------------------------------------------------------------*)
FC_DL_HexStringToBytes := 0;
nInvalidPos := 0;
uErrorId    := 16#0000_0000;
nBytes      := 0;

(*------------------------------------------------------------------------------
 * 段 2｜容量参数钳位：小于 1 抬到 1，大于 64 压到 64（瞬时码）
 *      Capacity clamp: raise to 1 or lower to 64, transient code
 *-----------------------------------------------------------------------------*)
IF nMaxBytes < 1 THEN
    nMaxBytes := 1;
    uErrorId  := 16#0001_0001;
ELSIF nMaxBytes > DL_HX_BUF_MAX THEN
    nMaxBytes := DL_HX_BUF_MAX;
    uErrorId  := 16#0001_0001;
END_IF

(*------------------------------------------------------------------------------
 * 段 3｜原文长度与有效区间初值（IEC 字符串位置 1 起）
 *      Original length and effective range init, IEC strings are 1-based
 *-----------------------------------------------------------------------------*)
nLen   := LEN(sHex);
nStart := 1;
nEnd   := nLen;

(*------------------------------------------------------------------------------
 * 段 4｜帧剥离（边界 B5）：只剥首冒号与尾部回车/换行，不剥空格。
 *      Framing strip: only the colon and trailing CR/LF, never spaces
 *      尾部先判换行再判回车，顺序固定，天然兼容 CRLF / LF / CR 三种结尾
 *-----------------------------------------------------------------------------*)
IF bStripFraming THEN
    IF (nLen >= 1) THEN
        sChar := MID(sHex, DL_HX_ONE, 1);
        IF sChar = DL_HX_COLON THEN
            nStart := 2;
        END_IF
    END_IF
    IF nEnd >= nStart THEN
        sChar := MID(sHex, DL_HX_ONE, nEnd);
        IF sChar = DL_HX_LF THEN
            nEnd := nEnd - 1;
        END_IF
    END_IF
    IF nEnd >= nStart THEN
        sChar := MID(sHex, DL_HX_ONE, nEnd);
        IF sChar = DL_HX_CR THEN
            nEnd := nEnd - 1;
        END_IF
    END_IF
END_IF

(*------------------------------------------------------------------------------
 * 段 5｜有效长度与空串兜底：空报文是合法输入，返回 0 不报错（边界 B7）
 *      Effective length and empty-string fallback: empty is legal, return 0
 *-----------------------------------------------------------------------------*)
nHexLen := nEnd - nStart + 1;
IF nHexLen < 0 THEN
    nHexLen := 0;
END_IF
IF nHexLen = 0 THEN
    RETURN;                                 // 空报文：返回 0、无故障 / Empty payload, return 0 with no error
END_IF

(*------------------------------------------------------------------------------
 * 段 6｜奇数长度拒绝（边界 B4）：判非法而非末尾补 0
 *      Odd length rejected: never pad a phantom byte
 *-----------------------------------------------------------------------------*)
IF (nHexLen MOD DL_HX_PAIR) <> 0 THEN
    uErrorId    := 16#0002_000A;            // 十六进制串非法 / Invalid hex string
    nInvalidPos := nStart + nHexLen;        // 指向悬空的半个字节 / Points at the dangling half byte
    FC_DL_HexStringToBytes := -1;
    RETURN;
END_IF

(*------------------------------------------------------------------------------
 * 段 7｜第一遍：全量字符合法性校验（标准 FIND 定位，大小写同等接受）
 *      Pass 1: full character validation via standard FIND, case-insensitive
 *      此遍绝不写输出缓冲（边界 B1）
 *-----------------------------------------------------------------------------*)
FOR nI := 0 TO (nHexLen - 1) DO
    sChar  := MID(sHex, DL_HX_ONE, nStart + nI);
    nHiNib := FIND(DL_HX_DIG_UP, sChar) - 1;    // 0..15，未命中为 -1 / 0..15, -1 if not found
    IF nHiNib < 0 THEN
        nHiNib := FIND(DL_HX_DIG_LOW, sChar) - 1;
    END_IF
    IF (nHiNib < 0) OR (nHiNib > 15) THEN
        uErrorId    := 16#0002_000A;        // 非 hex 字符 / Non-hex character
        nInvalidPos := nStart + nI;         // 原文 1 起位置（边界 B9） / 1-based original position
        FC_DL_HexStringToBytes := -1;
        RETURN;
    END_IF
END_FOR;

(*------------------------------------------------------------------------------
 * 段 8｜容量检查：整帧拒绝，不写半截（边界 B1）
 *      Capacity check: reject the whole frame, never write a partial stream
 *-----------------------------------------------------------------------------*)
nBytes := nHexLen / DL_HX_PAIR;             // 整除，奇数已在段 6 排除 / Integer division, odd already rejected
IF (nBytes > nMaxBytes) OR (nBytes > DL_HX_BUF_MAX) THEN
    uErrorId := 16#0001_0009;               // 输出缓冲不足 / Output buffer insufficient
    FC_DL_HexStringToBytes := -1;
    RETURN;
END_IF

(*------------------------------------------------------------------------------
 * 段 9｜第二遍：组装写入。高半字节左移 4 位或上低半字节，显式 INT_TO_BYTE
 *      Pass 2: assemble and write, explicit INT_TO_BYTE after the nibble shift
 *-----------------------------------------------------------------------------*)
FOR nI := 0 TO (nBytes - 1) DO
    sChar  := MID(sHex, DL_HX_ONE, nStart + (DL_HX_PAIR * nI));
    nHiNib := FIND(DL_HX_DIG_UP, sChar) - 1;
    IF nHiNib < 0 THEN
        nHiNib := FIND(DL_HX_DIG_LOW, sChar) - 1;
    END_IF
    sChar  := MID(sHex, DL_HX_ONE, nStart + (DL_HX_PAIR * nI) + 1);
    nLoNib := FIND(DL_HX_DIG_UP, sChar) - 1;
    IF nLoNib < 0 THEN
        nLoNib := FIND(DL_HX_DIG_LOW, sChar) - 1;
    END_IF
    IF (nI >= 0) AND (nI < DL_HX_BUF_MAX) THEN
        (* 写前下标双检（红线 R4）：容量已在段 8 保证，仍显式兜底 *)
        (* Index double check before writing: guaranteed by pass 8, explicit anyway *)
        aabyOut[nI] := SHL(INT_TO_BYTE(nHiNib), DL_HX_SHIFT) OR INT_TO_BYTE(nLoNib);
    END_IF
END_FOR;

(*------------------------------------------------------------------------------
 * 段 10｜成功返回：返回写入字节数；帧剥离发生时返回值不含帧字符
 *      Success return: byte count written, framing chars never counted
 *-----------------------------------------------------------------------------*)
FC_DL_HexStringToBytes := nBytes;
END_FUNCTION
